    IF NOT "FRK_PersistImages".D003.Rows[8].Used OR "FRK_PersistImages".D003.Rows[8].SchemaVersion <> 4 OR "FRK_PersistImages".D003.Rows[8].ModelCode <> 'MODEL_B' OR "FRK_PersistImages".D003.Rows[8].Record.Scope <> 'StationA.Cell.Gate' OR "FRK_PersistImages".D003.Rows[8].Record.WriteKey <> 'preset' OR "FRK_PersistImages".D003.Rows[8].Record.Revision <> 2 OR "FRK_PersistImages".D003.Rows[8].Record.Kind <> 0 OR "FRK_PersistImages".D003.Rows[8].Record.ValueType <> 0 THEN RETURN; END_IF;
    #Ok := "FRK_ConfigDecode"(Text := STRING_TO_WSTRING("FRK_PersistImages".D003.Rows[8].Record.ValueText), Storage := 3, Minimum := 0.0, Maximum := 1000.0, MaxLength := 0, Value := "FRK_ConfigScratch".Value);
    IF NOT #Ok THEN RETURN; END_IF;
    IF NOT "FRK_PersistImages".D003.Rows[9].Used OR "FRK_PersistImages".D003.Rows[9].SchemaVersion <> 4 OR "FRK_PersistImages".D003.Rows[9].ModelCode <> 'MODEL_B' OR "FRK_PersistImages".D003.Rows[9].Record.Scope <> 'StationA.Satellite' OR "FRK_PersistImages".D003.Rows[9].Record.WriteKey <> 'timeout' OR "FRK_PersistImages".D003.Rows[9].Record.Revision <> 1 OR "FRK_PersistImages".D003.Rows[9].Record.Kind <> 0 OR "FRK_PersistImages".D003.Rows[9].Record.ValueType <> 3 THEN RETURN; END_IF;
    #Ok := "FRK_ConfigDecode"(Text := STRING_TO_WSTRING("FRK_PersistImages".D003.Rows[9].Record.ValueText), Storage := 7, Minimum := 1.0, Maximum := 60000.0, MaxLength := 0, Value := "FRK_ConfigScratch".Value);
    IF NOT #Ok THEN RETURN; END_IF;
    IF NOT "FRK_PersistImages".D003.Rows[10].Used OR "FRK_PersistImages".D003.Rows[10].SchemaVersion <> 4 OR "FRK_PersistImages".D003.Rows[10].ModelCode <> 'MODEL_B' OR "FRK_PersistImages".D003.Rows[10].Record.Scope <> 'StationA.Satellite' OR "FRK_PersistImages".D003.Rows[10].Record.WriteKey <> 'preset' OR "FRK_PersistImages".D003.Rows[10].Record.Revision <> 2 OR "FRK_PersistImages".D003.Rows[10].Record.Kind <> 0 OR "FRK_PersistImages".D003.Rows[10].Record.ValueType <> 0 THEN RETURN; END_IF;
    #Ok := "FRK_ConfigDecode"(Text := STRING_TO_WSTRING("FRK_PersistImages".D003.Rows[10].Record.ValueText), Storage := 3, Minimum := 0.0, Maximum := 1000.0, MaxLength := 0, Value := "FRK_ConfigScratch".Value);
    IF NOT #Ok THEN RETURN; END_IF;
    IF NOT "FRK_PersistImages".D003.Rows[11].Used OR "FRK_PersistImages".D003.Rows[11].SchemaVersion <> 4 OR "FRK_PersistImages".D003.Rows[11].ModelCode <> 'MODEL_B' OR "FRK_PersistImages".D003.Rows[11].Record.Scope <> 'StationA.Satellite.Cell' OR "FRK_PersistImages".D003.Rows[11].Record.WriteKey <> 'timeout' OR "FRK_PersistImages".D003.Rows[11].Record.Revision <> 1 OR "FRK_PersistImages".D003.Rows[11].Record.Kind <> 0 OR "FRK_PersistImages".D003.Rows[11].Record.ValueType <> 3 THEN RETURN; END_IF;
    #Ok := "FRK_ConfigDecode"(Text := STRING_TO_WSTRING("FRK_PersistImages".D003.Rows[11].Record.ValueText), Storage := 7, Minimum := 1.0, Maximum := 60000.0, MaxLength := 0, Value := "FRK_ConfigScratch".Value);
    IF NOT #Ok THEN RETURN; END_IF;
    IF NOT "FRK_PersistImages".D003.Rows[12].Used OR "FRK_PersistImages".D003.Rows[12].SchemaVersion <> 4 OR "FRK_PersistImages".D003.Rows[12].ModelCode <> 'MODEL_B' OR "FRK_PersistImages".D003.Rows[12].Record.Scope <> 'StationA.Satellite.Cell' OR "FRK_PersistImages".D003.Rows[12].Record.WriteKey <> 'preset' OR "FRK_PersistImages".D003.Rows[12].Record.Revision <> 2 OR "FRK_PersistImages".D003.Rows[12].Record.Kind <> 0 OR "FRK_PersistImages".D003.Rows[12].Record.ValueType <> 0 THEN RETURN; END_IF;
    #Ok := "FRK_ConfigDecode"(Text := STRING_TO_WSTRING("FRK_PersistImages".D003.Rows[12].Record.ValueText), Storage := 3, Minimum := 0.0, Maximum := 1000.0, MaxLength := 0, Value := "FRK_ConfigScratch".Value);
    IF NOT #Ok THEN RETURN; END_IF;
    IF NOT "FRK_PersistImages".D003.Rows[13].Used OR "FRK_PersistImages".D003.Rows[13].SchemaVersion <> 4 OR "FRK_PersistImages".D003.Rows[13].ModelCode <> 'MODEL_B' OR "FRK_PersistImages".D003.Rows[13].Record.Scope <> 'StationA.Satellite.Cell.Clamp' OR "FRK_PersistImages".D003.Rows[13].Record.WriteKey <> 'timeout' OR "FRK_PersistImages".D003.Rows[13].Record.Revision <> 1 OR "FRK_PersistImages".D003.Rows[13].Record.Kind <> 0 OR "FRK_PersistImages".D003.Rows[13].Record.ValueType <> 3 THEN RETURN; END_IF;
    #Ok := "FRK_ConfigDecode"(Text := STRING_TO_WSTRING("FRK_PersistImages".D003.Rows[13].Record.ValueText), Storage := 7, Minimum := 1.0, Maximum := 60000.0, MaxLength := 0, Value := "FRK_ConfigScratch".Value);
    IF NOT #Ok THEN RETURN; END_IF;
    IF NOT "FRK_PersistImages".D003.Rows[14].Used OR "FRK_PersistImages".D003.Rows[14].SchemaVersion <> 4 OR "FRK_PersistImages".D003.Rows[14].ModelCode <> 'MODEL_B' OR "FRK_PersistImages".D003.Rows[14].Record.Scope <> 'StationA.Satellite.Cell.Clamp' OR "FRK_PersistImages".D003.Rows[14].Record.WriteKey <> 'preset' OR "FRK_PersistImages".D003.Rows[14].Record.Revision <> 2 OR "FRK_PersistImages".D003.Rows[14].Record.Kind <> 0 OR "FRK_PersistImages".D003.Rows[14].Record.ValueType <> 0 THEN RETURN; END_IF;
    #Ok := "FRK_ConfigDecode"(Text := STRING_TO_WSTRING("FRK_PersistImages".D003.Rows[14].Record.ValueText), Storage := 3, Minimum := 0.0, Maximum := 1000.0, MaxLength := 0, Value := "FRK_ConfigScratch".Value);
    IF NOT #Ok THEN RETURN; END_IF;
    IF NOT "FRK_PersistImages".D003.Rows[15].Used OR "FRK_PersistImages".D003.Rows[15].SchemaVersion <> 4 OR "FRK_PersistImages".D003.Rows[15].ModelCode <> 'MODEL_B' OR "FRK_PersistImages".D003.Rows[15].Record.Scope <> 'StationA.Satellite.Cell.Gate' OR "FRK_PersistImages".D003.Rows[15].Record.WriteKey <> 'timeout' OR "FRK_PersistImages".D003.Rows[15].Record.Revision <> 1 OR "FRK_PersistImages".D003.Rows[15].Record.Kind <> 0 OR "FRK_PersistImages".D003.Rows[15].Record.ValueType <> 3 THEN RETURN; END_IF;
    #Ok := "FRK_ConfigDecode"(Text := STRING_TO_WSTRING("FRK_PersistImages".D003.Rows[15].Record.ValueText), Storage := 7, Minimum := 1.0, Maximum := 60000.0, MaxLength := 0, Value := "FRK_ConfigScratch".Value);
    IF NOT #Ok THEN RETURN; END_IF;
    IF NOT "FRK_PersistImages".D003.Rows[16].Used OR "FRK_PersistImages".D003.Rows[16].SchemaVersion <> 4 OR "FRK_PersistImages".D003.Rows[16].ModelCode <> 'MODEL_B' OR "FRK_PersistImages".D003.Rows[16].Record.Scope <> 'StationA.Satellite.Cell.Gate' OR "FRK_PersistImages".D003.Rows[16].Record.WriteKey <> 'preset' OR "FRK_PersistImages".D003.Rows[16].Record.Revision <> 2 OR "FRK_PersistImages".D003.Rows[16].Record.Kind <> 0 OR "FRK_PersistImages".D003.Rows[16].Record.ValueType <> 0 THEN RETURN; END_IF;
    #Ok := "FRK_ConfigDecode"(Text := STRING_TO_WSTRING("FRK_PersistImages".D003.Rows[16].Record.ValueText), Storage := 3, Minimum := 0.0, Maximum := 1000.0, MaxLength := 0, Value := "FRK_ConfigScratch".Value);
    IF NOT #Ok THEN RETURN; END_IF;
    IF NOT "FRK_PersistImages".D003.Rows[17].Used OR "FRK_PersistImages".D003.Rows[17].SchemaVersion <> 4 OR "FRK_PersistImages".D003.Rows[17].ModelCode <> 'MODEL_B' OR "FRK_PersistImages".D003.Rows[17].Record.Scope <> 'StationA.Satellite.Inner' OR "FRK_PersistImages".D003.Rows[17].Record.WriteKey <> 'timeout' OR "FRK_PersistImages".D003.Rows[17].Record.Revision <> 1 OR "FRK_PersistImages".D003.Rows[17].Record.Kind <> 0 OR "FRK_PersistImages".D003.Rows[17].Record.ValueType <> 3 THEN RETURN; END_IF;
    #Ok := "FRK_ConfigDecode"(Text := STRING_TO_WSTRING("FRK_PersistImages".D003.Rows[17].Record.ValueText), Storage := 7, Minimum := 1.0, Maximum := 60000.0, MaxLength := 0, Value := "FRK_ConfigScratch".Value);
    IF NOT #Ok THEN RETURN; END_IF;
    IF NOT "FRK_PersistImages".D003.Rows[18].Used OR "FRK_PersistImages".D003.Rows[18].SchemaVersion <> 4 OR "FRK_PersistImages".D003.Rows[18].ModelCode <> 'MODEL_B' OR "FRK_PersistImages".D003.Rows[18].Record.Scope <> 'StationA.Satellite.Inner' OR "FRK_PersistImages".D003.Rows[18].Record.WriteKey <> 'preset' OR "FRK_PersistImages".D003.Rows[18].Record.Revision <> 2 OR "FRK_PersistImages".D003.Rows[18].Record.Kind <> 0 OR "FRK_PersistImages".D003.Rows[18].Record.ValueType <> 0 THEN RETURN; END_IF;
    #Ok := "FRK_ConfigDecode"(Text := STRING_TO_WSTRING("FRK_PersistImages".D003.Rows[18].Record.ValueText), Storage := 3, Minimum := 0.0, Maximum := 1000.0, MaxLength := 0, Value := "FRK_ConfigScratch".Value);
    IF NOT #Ok THEN RETURN; END_IF;
    IF NOT "FRK_PersistImages".D003.Rows[19].Used OR "FRK_PersistImages".D003.Rows[19].SchemaVersion <> 4 OR "FRK_PersistImages".D003.Rows[19].ModelCode <> 'MODEL_B' OR "FRK_PersistImages".D003.Rows[19].Record.Scope <> 'StationA.Satellite.Inner.Cell' OR "FRK_PersistImages".D003.Rows[19].Record.WriteKey <> 'timeout' OR "FRK_PersistImages".D003.Rows[19].Record.Revision <> 1 OR "FRK_PersistImages".D003.Rows[19].Record.Kind <> 0 OR "FRK_PersistImages".D003.Rows[19].Record.ValueType <> 3 THEN RETURN; END_IF;
    #Ok := "FRK_ConfigDecode"(Text := STRING_TO_WSTRING("FRK_PersistImages".D003.Rows[19].Record.ValueText), Storage := 7, Minimum := 1.0, Maximum := 60000.0, MaxLength := 0, Value := "FRK_ConfigScratch".Value);
    IF NOT #Ok THEN RETURN; END_IF;
    IF NOT "FRK_PersistImages".D003.Rows[20].Used OR "FRK_PersistImages".D003.Rows[20].SchemaVersion <> 4 OR "FRK_PersistImages".D003.Rows[20].ModelCode <> 'MODEL_B' OR "FRK_PersistImages".D003.Rows[20].Record.Scope <> 'StationA.Satellite.Inner.Cell' OR "FRK_PersistImages".D003.Rows[20].Record.WriteKey <> 'preset' OR "FRK_PersistImages".D003.Rows[20].Record.Revision <> 2 OR "FRK_PersistImages".D003.Rows[20].Record.Kind <> 0 OR "FRK_PersistImages".D003.Rows[20].Record.ValueType <> 0 THEN RETURN; END_IF;
    #Ok := "FRK_ConfigDecode"(Text := STRING_TO_WSTRING("FRK_PersistImages".D003.Rows[20].Record.ValueText), Storage := 3, Minimum := 0.0, Maximum := 1000.0, MaxLength := 0, Value := "FRK_ConfigScratch".Value);
    IF NOT #Ok THEN RETURN; END_IF;
    IF NOT "FRK_PersistImages".D003.Rows[21].Used OR "FRK_PersistImages".D003.Rows[21].SchemaVersion <> 4 OR "FRK_PersistImages".D003.Rows[21].ModelCode <> 'MODEL_B' OR "FRK_PersistImages".D003.Rows[21].Record.Scope <> 'StationA.Satellite.Inner.Cell.Clamp' OR "FRK_PersistImages".D003.Rows[21].Record.WriteKey <> 'timeout' OR "FRK_PersistImages".D003.Rows[21].Record.Revision <> 1 OR "FRK_PersistImages".D003.Rows[21].Record.Kind <> 0 OR "FRK_PersistImages".D003.Rows[21].Record.ValueType <> 3 THEN RETURN; END_IF;
    #Ok := "FRK_ConfigDecode"(Text := STRING_TO_WSTRING("FRK_PersistImages".D003.Rows[21].Record.ValueText), Storage := 7, Minimum := 1.0, Maximum := 60000.0, MaxLength := 0, Value := "FRK_ConfigScratch".Value);
    IF NOT #Ok THEN RETURN; END_IF;
    IF NOT "FRK_PersistImages".D003.Rows[22].Used OR "FRK_PersistImages".D003.Rows[22].SchemaVersion <> 4 OR "FRK_PersistImages".D003.Rows[22].ModelCode <> 'MODEL_B' OR "FRK_PersistImages".D003.Rows[22].Record.Scope <> 'StationA.Satellite.Inner.Cell.Clamp' OR "FRK_PersistImages".D003.Rows[22].Record.WriteKey <> 'preset' OR "FRK_PersistImages".D003.Rows[22].Record.Revision <> 2 OR "FRK_PersistImages".D003.Rows[22].Record.Kind <> 0 OR "FRK_PersistImages".D003.Rows[22].Record.ValueType <> 0 THEN RETURN; END_IF;
    #Ok := "FRK_ConfigDecode"(Text := STRING_TO_WSTRING("FRK_PersistImages".D003.Rows[22].Record.ValueText), Storage := 3, Minimum := 0.0, Maximum := 1000.0, MaxLength := 0, Value := "FRK_ConfigScratch".Value);
    IF NOT #Ok THEN RETURN; END_IF;
    IF NOT "FRK_PersistImages".D003.Rows[23].Used OR "FRK_PersistImages".D003.Rows[23].SchemaVersion <> 4 OR "FRK_PersistImages".D003.Rows[23].ModelCode <> 'MODEL_B' OR "FRK_PersistImages".D003.Rows[23].Record.Scope <> 'StationA.Satellite.Inner.Cell.Gate' OR "FRK_PersistImages".D003.Rows[23].Record.WriteKey <> 'timeout' OR "FRK_PersistImages".D003.Rows[23].Record.Revision <> 1 OR "FRK_PersistImages".D003.Rows[23].Record.Kind <> 0 OR "FRK_PersistImages".D003.Rows[23].Record.ValueType <> 3 THEN RETURN; END_IF;
    #Ok := "FRK_ConfigDecode"(Text := STRING_TO_WSTRING("FRK_PersistImages".D003.Rows[23].Record.ValueText), Storage := 7, Minimum := 1.0, Maximum := 60000.0, MaxLength := 0, Value := "FRK_ConfigScratch".Value);
    IF NOT #Ok THEN RETURN; END_IF;
    IF NOT "FRK_PersistImages".D003.Rows[24].Used OR "FRK_PersistImages".D003.Rows[24].SchemaVersion <> 4 OR "FRK_PersistImages".D003.Rows[24].ModelCode <> 'MODEL_B' OR "FRK_PersistImages".D003.Rows[24].Record.Scope <> 'StationA.Satellite.Inner.Cell.Gate' OR "FRK_PersistImages".D003.Rows[24].Record.WriteKey <> 'preset' OR "FRK_PersistImages".D003.Rows[24].Record.Revision <> 2 OR "FRK_PersistImages".D003.Rows[24].Record.Kind <> 0 OR "FRK_PersistImages".D003.Rows[24].Record.ValueType <> 0 THEN RETURN; END_IF;
    #Ok := "FRK_ConfigDecode"(Text := STRING_TO_WSTRING("FRK_PersistImages".D003.Rows[24].Record.ValueText), Storage := 3, Minimum := 0.0, Maximum := 1000.0, MaxLength := 0, Value := "FRK_ConfigScratch".Value);
    IF NOT #Ok THEN RETURN; END_IF;
    #Stored := "FRK_ConfigFind"(Scope := 'StationA', Key := 'timeout', ModelCode := 'MODEL_B');
    IF #Stored = 0 THEN
        FOR #Stored := 1 TO 108 DO IF NOT "FRK_ConfigStore".Rows[#Stored].Used THEN EXIT; END_IF; END_FOR;
    END_IF;
    IF #Stored < 1 OR #Stored > 108 THEN RETURN; END_IF;
    "FRK_ConfigStore".Rows[#Stored] := "FRK_PersistImages".D003.Rows[1];
    #Stored := "FRK_ConfigFind"(Scope := 'StationA', Key := 'preset', ModelCode := 'MODEL_B');
    IF #Stored = 0 THEN
        FOR #Stored := 1 TO 108 DO IF NOT "FRK_ConfigStore".Rows[#Stored].Used THEN EXIT; END_IF; END_FOR;
    END_IF;
    IF #Stored < 1 OR #Stored > 108 THEN RETURN; END_IF;
    "FRK_ConfigStore".Rows[#Stored] := "FRK_PersistImages".D003.Rows[2];
    #Stored := "FRK_ConfigFind"(Scope := 'StationA.Cell', Key := 'timeout', ModelCode := 'MODEL_B');
    IF #Stored = 0 THEN
        FOR #Stored := 1 TO 108 DO IF NOT "FRK_ConfigStore".Rows[#Stored].Used THEN EXIT; END_IF; END_FOR;
    END_IF;
    IF #Stored < 1 OR #Stored > 108 THEN RETURN; END_IF;
    "FRK_ConfigStore".Rows[#Stored] := "FRK_PersistImages".D003.Rows[3];
    #Stored := "FRK_ConfigFind"(Scope := 'StationA.Cell', Key := 'preset', ModelCode := 'MODEL_B');
    IF #Stored = 0 THEN
        FOR #Stored := 1 TO 108 DO IF NOT "FRK_ConfigStore".Rows[#Stored].Used THEN EXIT; END_IF; END_FOR;
    END_IF;
    IF #Stored < 1 OR #Stored > 108 THEN RETURN; END_IF;
    "FRK_ConfigStore".Rows[#Stored] := "FRK_PersistImages".D003.Rows[4];
    #Stored := "FRK_ConfigFind"(Scope := 'StationA.Cell.Clamp', Key := 'timeout', ModelCode := 'MODEL_B');
    IF #Stored = 0 THEN
        FOR #Stored := 1 TO 108 DO IF NOT "FRK_ConfigStore".Rows[#Stored].Used THEN EXIT; END_IF; END_FOR;
    END_IF;
    IF #Stored < 1 OR #Stored > 108 THEN RETURN; END_IF;
    "FRK_ConfigStore".Rows[#Stored] := "FRK_PersistImages".D003.Rows[5];
    #Stored := "FRK_ConfigFind"(Scope := 'StationA.Cell.Clamp', Key := 'preset', ModelCode := 'MODEL_B');
    IF #Stored = 0 THEN
        FOR #Stored := 1 TO 108 DO IF NOT "FRK_ConfigStore".Rows[#Stored].Used THEN EXIT; END_IF; END_FOR;
    END_IF;
    IF #Stored < 1 OR #Stored > 108 THEN RETURN; END_IF;
    "FRK_ConfigStore".Rows[#Stored] := "FRK_PersistImages".D003.Rows[6];
    #Stored := "FRK_ConfigFind"(Scope := 'StationA.Cell.Gate', Key := 'timeout', ModelCode := 'MODEL_B');
    IF #Stored = 0 THEN
        FOR #Stored := 1 TO 108 DO IF NOT "FRK_ConfigStore".Rows[#Stored].Used THEN EXIT; END_IF; END_FOR;
    END_IF;
    IF #Stored < 1 OR #Stored > 108 THEN RETURN; END_IF;
    "FRK_ConfigStore".Rows[#Stored] := "FRK_PersistImages".D003.Rows[7];
    #Stored := "FRK_ConfigFind"(Scope := 'StationA.Cell.Gate', Key := 'preset', ModelCode := 'MODEL_B');
    IF #Stored = 0 THEN
        FOR #Stored := 1 TO 108 DO IF NOT "FRK_ConfigStore".Rows[#Stored].Used THEN EXIT; END_IF; END_FOR;
    END_IF;
    IF #Stored < 1 OR #Stored > 108 THEN RETURN; END_IF;
    "FRK_ConfigStore".Rows[#Stored] := "FRK_PersistImages".D003.Rows[8];
    #Stored := "FRK_ConfigFind"(Scope := 'StationA.Satellite', Key := 'timeout', ModelCode := 'MODEL_B');
    IF #Stored = 0 THEN
        FOR #Stored := 1 TO 108 DO IF NOT "FRK_ConfigStore".Rows[#Stored].Used THEN EXIT; END_IF; END_FOR;
    END_IF;
    IF #Stored < 1 OR #Stored > 108 THEN RETURN; END_IF;
    "FRK_ConfigStore".Rows[#Stored] := "FRK_PersistImages".D003.Rows[9];
    #Stored := "FRK_ConfigFind"(Scope := 'StationA.Satellite', Key := 'preset', ModelCode := 'MODEL_B');
    IF #Stored = 0 THEN
        FOR #Stored := 1 TO 108 DO IF NOT "FRK_ConfigStore".Rows[#Stored].Used THEN EXIT; END_IF; END_FOR;
    END_IF;
    IF #Stored < 1 OR #Stored > 108 THEN RETURN; END_IF;
    "FRK_ConfigStore".Rows[#Stored] := "FRK_PersistImages".D003.Rows[10];
    #Stored := "FRK_ConfigFind"(Scope := 'StationA.Satellite.Cell', Key := 'timeout', ModelCode := 'MODEL_B');
    IF #Stored = 0 THEN
        FOR #Stored := 1 TO 108 DO IF NOT "FRK_ConfigStore".Rows[#Stored].Used THEN EXIT; END_IF; END_FOR;
    END_IF;
    IF #Stored < 1 OR #Stored > 108 THEN RETURN; END_IF;
    "FRK_ConfigStore".Rows[#Stored] := "FRK_PersistImages".D003.Rows[11];
    #Stored := "FRK_ConfigFind"(Scope := 'StationA.Satellite.Cell', Key := 'preset', ModelCode := 'MODEL_B');
    IF #Stored = 0 THEN
        FOR #Stored := 1 TO 108 DO IF NOT "FRK_ConfigStore".Rows[#Stored].Used THEN EXIT; END_IF; END_FOR;
    END_IF;
    IF #Stored < 1 OR #Stored > 108 THEN RETURN; END_IF;
    "FRK_ConfigStore".Rows[#Stored] := "FRK_PersistImages".D003.Rows[12];
    #Stored := "FRK_ConfigFind"(Scope := 'StationA.Satellite.Cell.Clamp', Key := 'timeout', ModelCode := 'MODEL_B');
    IF #Stored = 0 THEN
        FOR #Stored := 1 TO 108 DO IF NOT "FRK_ConfigStore".Rows[#Stored].Used THEN EXIT; END_IF; END_FOR;
    END_IF;
    IF #Stored < 1 OR #Stored > 108 THEN RETURN; END_IF;
    "FRK_ConfigStore".Rows[#Stored] := "FRK_PersistImages".D003.Rows[13];
    #Stored := "FRK_ConfigFind"(Scope := 'StationA.Satellite.Cell.Clamp', Key := 'preset', ModelCode := 'MODEL_B');
    IF #Stored = 0 THEN
        FOR #Stored := 1 TO 108 DO IF NOT "FRK_ConfigStore".Rows[#Stored].Used THEN EXIT; END_IF; END_FOR;
    END_IF;
    IF #Stored < 1 OR #Stored > 108 THEN RETURN; END_IF;
    "FRK_ConfigStore".Rows[#Stored] := "FRK_PersistImages".D003.Rows[14];
    #Stored := "FRK_ConfigFind"(Scope := 'StationA.Satellite.Cell.Gate', Key := 'timeout', ModelCode := 'MODEL_B');
    IF #Stored = 0 THEN
        FOR #Stored := 1 TO 108 DO IF NOT "FRK_ConfigStore".Rows[#Stored].Used THEN EXIT; END_IF; END_FOR;
    END_IF;
    IF #Stored < 1 OR #Stored > 108 THEN RETURN; END_IF;
    "FRK_ConfigStore".Rows[#Stored] := "FRK_PersistImages".D003.Rows[15];
    #Stored := "FRK_ConfigFind"(Scope := 'StationA.Satellite.Cell.Gate', Key := 'preset', ModelCode := 'MODEL_B');
    IF #Stored = 0 THEN
        FOR #Stored := 1 TO 108 DO IF NOT "FRK_ConfigStore".Rows[#Stored].Used THEN EXIT; END_IF; END_FOR;
    END_IF;
    IF #Stored < 1 OR #Stored > 108 THEN RETURN; END_IF;
    "FRK_ConfigStore".Rows[#Stored] := "FRK_PersistImages".D003.Rows[16];
    #Stored := "FRK_ConfigFind"(Scope := 'StationA.Satellite.Inner', Key := 'timeout', ModelCode := 'MODEL_B');
    IF #Stored = 0 THEN
        FOR #Stored := 1 TO 108 DO IF NOT "FRK_ConfigStore".Rows[#Stored].Used THEN EXIT; END_IF; END_FOR;
    END_IF;
    IF #Stored < 1 OR #Stored > 108 THEN RETURN; END_IF;
    "FRK_ConfigStore".Rows[#Stored] := "FRK_PersistImages".D003.Rows[17];
    #Stored := "FRK_ConfigFind"(Scope := 'StationA.Satellite.Inner', Key := 'preset', ModelCode := 'MODEL_B');
    IF #Stored = 0 THEN
        FOR #Stored := 1 TO 108 DO IF NOT "FRK_ConfigStore".Rows[#Stored].Used THEN EXIT; END_IF; END_FOR;
    END_IF;
    IF #Stored < 1 OR #Stored > 108 THEN RETURN; END_IF;
    "FRK_ConfigStore".Rows[#Stored] := "FRK_PersistImages".D003.Rows[18];
    #Stored := "FRK_ConfigFind"(Scope := 'StationA.Satellite.Inner.Cell', Key := 'timeout', ModelCode := 'MODEL_B');
    IF #Stored = 0 THEN
        FOR #Stored := 1 TO 108 DO IF NOT "FRK_ConfigStore".Rows[#Stored].Used THEN EXIT; END_IF; END_FOR;
    END_IF;
    IF #Stored < 1 OR #Stored > 108 THEN RETURN; END_IF;
    "FRK_ConfigStore".Rows[#Stored] := "FRK_PersistImages".D003.Rows[19];
    #Stored := "FRK_ConfigFind"(Scope := 'StationA.Satellite.Inner.Cell', Key := 'preset', ModelCode := 'MODEL_B');
    IF #Stored = 0 THEN
        FOR #Stored := 1 TO 108 DO IF NOT "FRK_ConfigStore".Rows[#Stored].Used THEN EXIT; END_IF; END_FOR;
    END_IF;
    IF #Stored < 1 OR #Stored > 108 THEN RETURN; END_IF;
    "FRK_ConfigStore".Rows[#Stored] := "FRK_PersistImages".D003.Rows[20];
    #Stored := "FRK_ConfigFind"(Scope := 'StationA.Satellite.Inner.Cell.Clamp', Key := 'timeout', ModelCode := 'MODEL_B');
    IF #Stored = 0 THEN
        FOR #Stored := 1 TO 108 DO IF NOT "FRK_ConfigStore".Rows[#Stored].Used THEN EXIT; END_IF; END_FOR;
    END_IF;
    IF #Stored < 1 OR #Stored > 108 THEN RETURN; END_IF;
    "FRK_ConfigStore".Rows[#Stored] := "FRK_PersistImages".D003.Rows[21];
    #Stored := "FRK_ConfigFind"(Scope := 'StationA.Satellite.Inner.Cell.Clamp', Key := 'preset', ModelCode := 'MODEL_B');
    IF #Stored = 0 THEN
        FOR #Stored := 1 TO 108 DO IF NOT "FRK_ConfigStore".Rows[#Stored].Used THEN EXIT; END_IF; END_FOR;
    END_IF;
    IF #Stored < 1 OR #Stored > 108 THEN RETURN; END_IF;
    "FRK_ConfigStore".Rows[#Stored] := "FRK_PersistImages".D003.Rows[22];
    #Stored := "FRK_ConfigFind"(Scope := 'StationA.Satellite.Inner.Cell.Gate', Key := 'timeout', ModelCode := 'MODEL_B');
    IF #Stored = 0 THEN
        FOR #Stored := 1 TO 108 DO IF NOT "FRK_ConfigStore".Rows[#Stored].Used THEN EXIT; END_IF; END_FOR;
    END_IF;
    IF #Stored < 1 OR #Stored > 108 THEN RETURN; END_IF;
    "FRK_ConfigStore".Rows[#Stored] := "FRK_PersistImages".D003.Rows[23];
    #Stored := "FRK_ConfigFind"(Scope := 'StationA.Satellite.Inner.Cell.Gate', Key := 'preset', ModelCode := 'MODEL_B');
    IF #Stored = 0 THEN
        FOR #Stored := 1 TO 108 DO IF NOT "FRK_ConfigStore".Rows[#Stored].Used THEN EXIT; END_IF; END_FOR;
    END_IF;
    IF #Stored < 1 OR #Stored > 108 THEN RETURN; END_IF;
    "FRK_ConfigStore".Rows[#Stored] := "FRK_PersistImages".D003.Rows[24];
    "FRK_ConfigStore".SchemaVersion := 1;
    #FRK_DocApply_D003 := TRUE;
END_FUNCTION
FUNCTION "FRK_DocCapture_D004" : Bool
{ S7_Optimized_Access := 'TRUE' }
VERSION : 0.1
VAR_IN_OUT
    Length : DInt;
END_VAR
VAR_TEMP
    Index : Int;
    Stored : Int;
    Position : DInt;
    NativeResult : Int;
    Ok : Bool;
END_VAR
BEGIN
    #FRK_DocCapture_D004 := FALSE;
    "FRK_PersistImages".D004.SchemaVersion := 1; "FRK_PersistImages".D004.Scope := 'StationA';
    #Stored := 0;
    FOR #Index := 1 TO 2 DO
        IF "FRK_AccessPolicies".Rows[#Index].Scope = 'StationA' THEN #Stored := #Index; END_IF;
    END_FOR;
    IF #Stored = 0 THEN RETURN; END_IF;
    "FRK_PersistImages".D004.Image := "FRK_AccessPolicies".Rows[#Stored];
    IF NOT "FRK_AccessPolicyValid"(Image := "FRK_PersistImages".D004.Image) THEN RETURN; END_IF;
    FOR #Index := 0 TO 413 DO "FRK_PersistBuffers".D004Data[#Index] := BYTE#0; END_FOR;
    #Position := 24;
    #NativeResult := Serialize(SRC_VARIABLE := "FRK_PersistImages".D004, DEST_ARRAY => "FRK_PersistBuffers".D004Data, POS := #Position);
    IF #NativeResult <> 0 OR #Position < 24 OR #Position > 414 THEN RETURN; END_IF;
    #Length := #Position - 24;
    #FRK_DocCapture_D004 := TRUE;
END_FUNCTION
FUNCTION "FRK_DocApply_D004" : Bool
{ S7_Optimized_Access := 'TRUE' }
VERSION : 0.1
VAR_TEMP
    Index : Int;
    Stored : Int;
    Position : DInt;
    NativeResult : Int;
    Ok : Bool;
END_VAR
BEGIN
    #FRK_DocApply_D004 := FALSE;
    #Position := 24;
    #NativeResult := Deserialize(SRC_ARRAY := "FRK_PersistBuffers".D004Data, DEST_VARIABLE => "FRK_PersistImages".D004, POS := #Position);
    IF #NativeResult <> 0 OR #Position <> 24 + UDINT_TO_DINT("FRK_PersistConsumers".Rows[4].Result.Length) THEN RETURN; END_IF;
    IF "FRK_PersistImages".D004.SchemaVersion <> 1 OR "FRK_PersistImages".D004.Scope <> 'StationA' THEN RETURN; END_IF;
    IF "FRK_PersistImages".D004.Image.Scope <> 'StationA' OR NOT "FRK_AccessPolicyValid"(Image := "FRK_PersistImages".D004.Image) THEN RETURN; END_IF;
    "FRK_AccessPolicies".Rows[1] := "FRK_PersistImages".D004.Image;
    #FRK_DocApply_D004 := TRUE;
END_FUNCTION
FUNCTION "FRK_DocCapture_D005" : Bool
{ S7_Optimized_Access := 'TRUE' }
VERSION : 0.1
VAR_IN_OUT
    Length : DInt;
END_VAR
VAR_TEMP
    Index : Int;
    Stored : Int;
    Position : DInt;
    NativeResult : Int;
    Ok : Bool;
END_VAR
BEGIN
    #FRK_DocCapture_D005 := FALSE;
    "FRK_PersistImages".D005.SchemaVersion := 1; "FRK_PersistImages".D005.Scope := 'StationB';
    "FRK_PersistImages".D005.Kind := 1;
    "FRK_PersistImages".D005.ModelCode := '';
    "FRK_PersistImages".D005.ActiveModel := "FRK_ConfigStore".ActiveModels[2];
    "FRK_PersistImages".D005.Count := 6;
    #Stored := "FRK_ConfigFind"(Scope := 'StationB', Key := 'siteLabel', ModelCode := '');
    IF #Stored = 0 THEN RETURN; END_IF;
    "FRK_PersistImages".D005.Rows[1] := "FRK_ConfigStore".Rows[#Stored];
    #Stored := "FRK_ConfigFind"(Scope := 'StationB', Key := 'enabled', ModelCode := '');
    IF #Stored = 0 THEN RETURN; END_IF;
    "FRK_PersistImages".D005.Rows[2] := "FRK_ConfigStore".Rows[#Stored];
    #Stored := "FRK_ConfigFind"(Scope := 'StationB.Satellite', Key := 'siteLabel', ModelCode := '');
    IF #Stored = 0 THEN RETURN; END_IF;
    "FRK_PersistImages".D005.Rows[3] := "FRK_ConfigStore".Rows[#Stored];
    #Stored := "FRK_ConfigFind"(Scope := 'StationB.Satellite', Key := 'enabled', ModelCode := '');
    IF #Stored = 0 THEN RETURN; END_IF;
    "FRK_PersistImages".D005.Rows[4] := "FRK_ConfigStore".Rows[#Stored];
    #Stored := "FRK_ConfigFind"(Scope := 'StationB.Satellite.Inner', Key := 'siteLabel', ModelCode := '');
    IF #Stored = 0 THEN RETURN; END_IF;
    "FRK_PersistImages".D005.Rows[5] := "FRK_ConfigStore".Rows[#Stored];
    #Stored := "FRK_ConfigFind"(Scope := 'StationB.Satellite.Inner', Key := 'enabled', ModelCode := '');
    IF #Stored = 0 THEN RETURN; END_IF;
    "FRK_PersistImages".D005.Rows[6] := "FRK_ConfigStore".Rows[#Stored];
    FOR #Index := 0 TO 3085 DO "FRK_PersistBuffers".D005Data[#Index] := BYTE#0; END_FOR;
    #Position := 24;
    #NativeResult := Serialize(SRC_VARIABLE := "FRK_PersistImages".D005, DEST_ARRAY => "FRK_PersistBuffers".D005Data, POS := #Position);
    IF #NativeResult <> 0 OR #Position < 24 OR #Position > 3086 THEN RETURN; END_IF;
    #Length := #Position - 24;
    #FRK_DocCapture_D005 := TRUE;
END_FUNCTION
FUNCTION "FRK_DocApply_D005" : Bool
{ S7_Optimized_Access := 'TRUE' }
VERSION : 0.1
VAR_TEMP
    Index : Int;
    Stored : Int;
    Position : DInt;
    NativeResult : Int;
    Ok : Bool;
END_VAR
BEGIN
    #FRK_DocApply_D005 := FALSE;
    #Position := 24;
    #NativeResult := Deserialize(SRC_ARRAY := "FRK_PersistBuffers".D005Data, DEST_VARIABLE => "FRK_PersistImages".D005, POS := #Position);
    IF #NativeResult <> 0 OR #Position <> 24 + UDINT_TO_DINT("FRK_PersistConsumers".Rows[5].Result.Length) THEN RETURN; END_IF;
    IF "FRK_PersistImages".D005.SchemaVersion <> 1 OR "FRK_PersistImages".D005.Scope <> 'StationB' THEN RETURN; END_IF;
    IF "FRK_PersistImages".D005.Kind <> 1 OR "FRK_PersistImages".D005.ModelCode <> '' OR "FRK_PersistImages".D005.Count <> 6 THEN RETURN; END_IF;
    IF "FRK_PersistImages".D005.ActiveModel <> 'MODEL_A' AND "FRK_PersistImages".D005.ActiveModel <> 'MODEL_B' THEN RETURN; END_IF;
    IF NOT "FRK_PersistImages".D005.Rows[1].Used OR "FRK_PersistImages".D005.Rows[1].SchemaVersion <> 1 OR "FRK_PersistImages".D005.Rows[1].ModelCode <> '' OR "FRK_PersistImages".D005.Rows[1].Record.Scope <> 'StationB' OR "FRK_PersistImages".D005.Rows[1].Record.WriteKey <> 'siteLabel' OR "FRK_PersistImages".D005.Rows[1].Record.Revision <> 1 OR "FRK_PersistImages".D005.Rows[1].Record.Kind <> 1 OR "FRK_PersistImages".D005.Rows[1].Record.ValueType <> 1 THEN RETURN; END_IF;
    #Ok := "FRK_ConfigDecode"(Text := STRING_TO_WSTRING("FRK_PersistImages".D005.Rows[1].Record.ValueText), Storage := 8, Minimum := 0.0, Maximum := 1.0, MaxLength := 80, Value := "FRK_ConfigScratch".Value);
    IF NOT #Ok THEN RETURN; END_IF;
    IF NOT "FRK_PersistImages".D005.Rows[2].Used OR "FRK_PersistImages".D005.Rows[2].SchemaVersion <> 1 OR "FRK_PersistImages".D005.Rows[2].ModelCode <> '' OR "FRK_PersistImages".D005.Rows[2].Record.Scope <> 'StationB' OR "FRK_PersistImages".D005.Rows[2].Record.WriteKey <> 'enabled' OR "FRK_PersistImages".D005.Rows[2].Record.Revision <> 1 OR "FRK_PersistImages".D005.Rows[2].Record.Kind <> 1 OR "FRK_PersistImages".D005.Rows[2].Record.ValueType <> 2 THEN RETURN; END_IF;
    #Ok := "FRK_ConfigDecode"(Text := STRING_TO_WSTRING("FRK_PersistImages".D005.Rows[2].Record.ValueText), Storage := 1, Minimum := 0.0, Maximum := 1.0, MaxLength := 0, Value := "FRK_ConfigScratch".Value);
    IF NOT #Ok THEN RETURN; END_IF;
    IF NOT "FRK_PersistImages".D005.Rows[3].Used OR "FRK_PersistImages".D005.Rows[3].SchemaVersion <> 1 OR "FRK_PersistImages".D005.Rows[3].ModelCode <> '' OR "FRK_PersistImages".D005.Rows[3].Record.Scope <> 'StationB.Satellite' OR "FRK_PersistImages".D005.Rows[3].Record.WriteKey <> 'siteLabel' OR "FRK_PersistImages".D005.Rows[3].Record.Revision <> 1 OR "FRK_PersistImages".D005.Rows[3].Record.Kind <> 1 OR "FRK_PersistImages".D005.Rows[3].Record.ValueType <> 1 THEN RETURN; END_IF;
    #Ok := "FRK_ConfigDecode"(Text := STRING_TO_WSTRING("FRK_PersistImages".D005.Rows[3].Record.ValueText), Storage := 8, Minimum := 0.0, Maximum := 1.0, MaxLength := 80, Value := "FRK_ConfigScratch".Value);
    IF NOT #Ok THEN RETURN; END_IF;
    IF NOT "FRK_PersistImages".D005.Rows[4].Used OR "FRK_PersistImages".D005.Rows[4].SchemaVersion <> 1 OR "FRK_PersistImages".D005.Rows[4].ModelCode <> '' OR "FRK_PersistImages".D005.Rows[4].Record.Scope <> 'StationB.Satellite' OR "FRK_PersistImages".D005.Rows[4].Record.WriteKey <> 'enabled' OR "FRK_PersistImages".D005.Rows[4].Record.Revision <> 1 OR "FRK_PersistImages".D005.Rows[4].Record.Kind <> 1 OR "FRK_PersistImages".D005.Rows[4].Record.ValueType <> 2 THEN RETURN; END_IF;
    #Ok := "FRK_ConfigDecode"(Text := STRING_TO_WSTRING("FRK_PersistImages".D005.Rows[4].Record.ValueText), Storage := 1, Minimum := 0.0, Maximum := 1.0, MaxLength := 0, Value := "FRK_ConfigScratch".Value);
    IF NOT #Ok THEN RETURN; END_IF;
    IF NOT "FRK_PersistImages".D005.Rows[5].Used OR "FRK_PersistImages".D005.Rows[5].SchemaVersion <> 1 OR "FRK_PersistImages".D005.Rows[5].ModelCode <> '' OR "FRK_PersistImages".D005.Rows[5].Record.Scope <> 'StationB.Satellite.Inner' OR "FRK_PersistImages".D005.Rows[5].Record.WriteKey <> 'siteLabel' OR "FRK_PersistImages".D005.Rows[5].Record.Revision <> 1 OR "FRK_PersistImages".D005.Rows[5].Record.Kind <> 1 OR "FRK_PersistImages".D005.Rows[5].Record.ValueType <> 1 THEN RETURN; END_IF;
    #Ok := "FRK_ConfigDecode"(Text := STRING_TO_WSTRING("FRK_PersistImages".D005.Rows[5].Record.ValueText), Storage := 8, Minimum := 0.0, Maximum := 1.0, MaxLength := 80, Value := "FRK_ConfigScratch".Value);
    IF NOT #Ok THEN RETURN; END_IF;
    IF NOT "FRK_PersistImages".D005.Rows[6].Used OR "FRK_PersistImages".D005.Rows[6].SchemaVersion <> 1 OR "FRK_PersistImages".D005.Rows[6].ModelCode <> '' OR "FRK_PersistImages".D005.Rows[6].Record.Scope <> 'StationB.Satellite.Inner' OR "FRK_PersistImages".D005.Rows[6].Record.WriteKey <> 'enabled' OR "FRK_PersistImages".D005.Rows[6].Record.Revision <> 1 OR "FRK_PersistImages".D005.Rows[6].Record.Kind <> 1 OR "FRK_PersistImages".D005.Rows[6].Record.ValueType <> 2 THEN RETURN; END_IF;
    #Ok := "FRK_ConfigDecode"(Text := STRING_TO_WSTRING("FRK_PersistImages".D005.Rows[6].Record.ValueText), Storage := 1, Minimum := 0.0, Maximum := 1.0, MaxLength := 0, Value := "FRK_ConfigScratch".Value);
    IF NOT #Ok THEN RETURN; END_IF;
    #Stored := "FRK_ConfigFind"(Scope := 'StationB', Key := 'siteLabel', ModelCode := '');
    IF #Stored = 0 THEN
        FOR #Stored := 1 TO 108 DO IF NOT "FRK_ConfigStore".Rows[#Stored].Used THEN EXIT; END_IF; END_FOR;
    END_IF;
    IF #Stored < 1 OR #Stored > 108 THEN RETURN; END_IF;
    "FRK_ConfigStore".Rows[#Stored] := "FRK_PersistImages".D005.Rows[1];
    #Stored := "FRK_ConfigFind"(Scope := 'StationB', Key := 'enabled', ModelCode := '');
    IF #Stored = 0 THEN
        FOR #Stored := 1 TO 108 DO IF NOT "FRK_ConfigStore".Rows[#Stored].Used THEN EXIT; END_IF; END_FOR;
    END_IF;
    IF #Stored < 1 OR #Stored > 108 THEN RETURN; END_IF;
    "FRK_ConfigStore".Rows[#Stored] := "FRK_PersistImages".D005.Rows[2];
    #Stored := "FRK_ConfigFind"(Scope := 'StationB.Satellite', Key := 'siteLabel', ModelCode := '');
    IF #Stored = 0 THEN
        FOR #Stored := 1 TO 108 DO IF NOT "FRK_ConfigStore".Rows[#Stored].Used THEN EXIT; END_IF; END_FOR;
    END_IF;
    IF #Stored < 1 OR #Stored > 108 THEN RETURN; END_IF;
    "FRK_ConfigStore".Rows[#Stored] := "FRK_PersistImages".D005.Rows[3];
    #Stored := "FRK_ConfigFind"(Scope := 'StationB.Satellite', Key := 'enabled', ModelCode := '');
    IF #Stored = 0 THEN
        FOR #Stored := 1 TO 108 DO IF NOT "FRK_ConfigStore".Rows[#Stored].Used THEN EXIT; END_IF; END_FOR;
    END_IF;
    IF #Stored < 1 OR #Stored > 108 THEN RETURN; END_IF;
    "FRK_ConfigStore".Rows[#Stored] := "FRK_PersistImages".D005.Rows[4];
    #Stored := "FRK_ConfigFind"(Scope := 'StationB.Satellite.Inner', Key := 'siteLabel', ModelCode := '');
    IF #Stored = 0 THEN
        FOR #Stored := 1 TO 108 DO IF NOT "FRK_ConfigStore".Rows[#Stored].Used THEN EXIT; END_IF; END_FOR;
    END_IF;
    IF #Stored < 1 OR #Stored > 108 THEN RETURN; END_IF;
    "FRK_ConfigStore".Rows[#Stored] := "FRK_PersistImages".D005.Rows[5];
    #Stored := "FRK_ConfigFind"(Scope := 'StationB.Satellite.Inner', Key := 'enabled', ModelCode := '');
    IF #Stored = 0 THEN
        FOR #Stored := 1 TO 108 DO IF NOT "FRK_ConfigStore".Rows[#Stored].Used THEN EXIT; END_IF; END_FOR;
    END_IF;
    IF #Stored < 1 OR #Stored > 108 THEN RETURN; END_IF;
    "FRK_ConfigStore".Rows[#Stored] := "FRK_PersistImages".D005.Rows[6];
    "FRK_ConfigStore".ActiveModels[2] := "FRK_PersistImages".D005.ActiveModel;
    "FRK_ConfigStore".SchemaVersion := 1;
    #FRK_DocApply_D005 := TRUE;
END_FUNCTION
FUNCTION "FRK_DocCapture_D006" : Bool
{ S7_Optimized_Access := 'TRUE' }
VERSION : 0.1
VAR_IN_OUT
    Length : DInt;
END_VAR
VAR_TEMP
    Index : Int;
    Stored : Int;
    Position : DInt;
    NativeResult : Int;
    Ok : Bool;
END_VAR
BEGIN
    #FRK_DocCapture_D006 := FALSE;
    "FRK_PersistImages".D006.SchemaVersion := 1; "FRK_PersistImages".D006.Scope := 'StationB';
    "FRK_PersistImages".D006.Kind := 0;
    "FRK_PersistImages".D006.ModelCode := 'MODEL_A';
    "FRK_PersistImages".D006.ActiveModel := "FRK_ConfigStore".ActiveModels[2];
    "FRK_PersistImages".D006.Count := 24;
    #Stored := "FRK_ConfigFind"(Scope := 'StationB', Key := 'timeout', ModelCode := 'MODEL_A');
    IF #Stored = 0 THEN RETURN; END_IF;
    "FRK_PersistImages".D006.Rows[1] := "FRK_ConfigStore".Rows[#Stored];
    #Stored := "FRK_ConfigFind"(Scope := 'StationB', Key := 'preset', ModelCode := 'MODEL_A');
    IF #Stored = 0 THEN RETURN; END_IF;
    "FRK_PersistImages".D006.Rows[2] := "FRK_ConfigStore".Rows[#Stored];
    #Stored := "FRK_ConfigFind"(Scope := 'StationB.Cell', Key := 'timeout', ModelCode := 'MODEL_A');
    IF #Stored = 0 THEN RETURN; END_IF;
    "FRK_PersistImages".D006.Rows[3] := "FRK_ConfigStore".Rows[#Stored];
    #Stored := "FRK_ConfigFind"(Scope := 'StationB.Cell', Key := 'preset', ModelCode := 'MODEL_A');
    IF #Stored = 0 THEN RETURN; END_IF;
    "FRK_PersistImages".D006.Rows[4] := "FRK_ConfigStore".Rows[#Stored];
    #Stored := "FRK_ConfigFind"(Scope := 'StationB.Cell.Clamp', Key := 'timeout', ModelCode := 'MODEL_A');
    IF #Stored = 0 THEN RETURN; END_IF;
    "FRK_PersistImages".D006.Rows[5] := "FRK_ConfigStore".Rows[#Stored];
    #Stored := "FRK_ConfigFind"(Scope := 'StationB.Cell.Clamp', Key := 'preset', ModelCode := 'MODEL_A');
    IF #Stored = 0 THEN RETURN; END_IF;
    "FRK_PersistImages".D006.Rows[6] := "FRK_ConfigStore".Rows[#Stored];
    #Stored := "FRK_ConfigFind"(Scope := 'StationB.Cell.Gate', Key := 'timeout', ModelCode := 'MODEL_A');
    IF #Stored = 0 THEN RETURN; END_IF;
    "FRK_PersistImages".D006.Rows[7] := "FRK_ConfigStore".Rows[#Stored];
    #Stored := "FRK_ConfigFind"(Scope := 'StationB.Cell.Gate', Key := 'preset', ModelCode := 'MODEL_A');
    IF #Stored = 0 THEN RETURN; END_IF;
    "FRK_PersistImages".D006.Rows[8] := "FRK_ConfigStore".Rows[#Stored];
    #Stored := "FRK_ConfigFind"(Scope := 'StationB.Satellite', Key := 'timeout', ModelCode := 'MODEL_A');
    IF #Stored = 0 THEN RETURN; END_IF;
    "FRK_PersistImages".D006.Rows[9] := "FRK_ConfigStore".Rows[#Stored];
    #Stored := "FRK_ConfigFind"(Scope := 'StationB.Satellite', Key := 'preset', ModelCode := 'MODEL_A');
    IF #Stored = 0 THEN RETURN; END_IF;
    "FRK_PersistImages".D006.Rows[10] := "FRK_ConfigStore".Rows[#Stored];
    #Stored := "FRK_ConfigFind"(Scope := 'StationB.Satellite.Cell', Key := 'timeout', ModelCode := 'MODEL_A');
    IF #Stored = 0 THEN RETURN; END_IF;
    "FRK_PersistImages".D006.Rows[11] := "FRK_ConfigStore".Rows[#Stored];
    #Stored := "FRK_ConfigFind"(Scope := 'StationB.Satellite.Cell', Key := 'preset', ModelCode := 'MODEL_A');
    IF #Stored = 0 THEN RETURN; END_IF;
    "FRK_PersistImages".D006.Rows[12] := "FRK_ConfigStore".Rows[#Stored];
    #Stored := "FRK_ConfigFind"(Scope := 'StationB.Satellite.Cell.Clamp', Key := 'timeout', ModelCode := 'MODEL_A');
    IF #Stored = 0 THEN RETURN; END_IF;
    "FRK_PersistImages".D006.Rows[13] := "FRK_ConfigStore".Rows[#Stored];
    #Stored := "FRK_ConfigFind"(Scope := 'StationB.Satellite.Cell.Clamp', Key := 'preset', ModelCode := 'MODEL_A');
    IF #Stored = 0 THEN RETURN; END_IF;
    "FRK_PersistImages".D006.Rows[14] := "FRK_ConfigStore".Rows[#Stored];
    #Stored := "FRK_ConfigFind"(Scope := 'StationB.Satellite.Cell.Gate', Key := 'timeout', ModelCode := 'MODEL_A');
    IF #Stored = 0 THEN RETURN; END_IF;
    "FRK_PersistImages".D006.Rows[15] := "FRK_ConfigStore".Rows[#Stored];
    #Stored := "FRK_ConfigFind"(Scope := 'StationB.Satellite.Cell.Gate', Key := 'preset', ModelCode := 'MODEL_A');
    IF #Stored = 0 THEN RETURN; END_IF;
    "FRK_PersistImages".D006.Rows[16] := "FRK_ConfigStore".Rows[#Stored];
    #Stored := "FRK_ConfigFind"(Scope := 'StationB.Satellite.Inner', Key := 'timeout', ModelCode := 'MODEL_A');
    IF #Stored = 0 THEN RETURN; END_IF;
    "FRK_PersistImages".D006.Rows[17] := "FRK_ConfigStore".Rows[#Stored];
    #Stored := "FRK_ConfigFind"(Scope := 'StationB.Satellite.Inner', Key := 'preset', ModelCode := 'MODEL_A');
    IF #Stored = 0 THEN RETURN; END_IF;
    "FRK_PersistImages".D006.Rows[18] := "FRK_ConfigStore".Rows[#Stored];
    #Stored := "FRK_ConfigFind"(Scope := 'StationB.Satellite.Inner.Cell', Key := 'timeout', ModelCode := 'MODEL_A');
    IF #Stored = 0 THEN RETURN; END_IF;
    "FRK_PersistImages".D006.Rows[19] := "FRK_ConfigStore".Rows[#Stored];
    #Stored := "FRK_ConfigFind"(Scope := 'StationB.Satellite.Inner.Cell', Key := 'preset', ModelCode := 'MODEL_A');
    IF #Stored = 0 THEN RETURN; END_IF;
    "FRK_PersistImages".D006.Rows[20] := "FRK_ConfigStore".Rows[#Stored];
    #Stored := "FRK_ConfigFind"(Scope := 'StationB.Satellite.Inner.Cell.Clamp', Key := 'timeout', ModelCode := 'MODEL_A');
    IF #Stored = 0 THEN RETURN; END_IF;
    "FRK_PersistImages".D006.Rows[21] := "FRK_ConfigStore".Rows[#Stored];
    #Stored := "FRK_ConfigFind"(Scope := 'StationB.Satellite.Inner.Cell.Clamp', Key := 'preset', ModelCode := 'MODEL_A');
    IF #Stored = 0 THEN RETURN; END_IF;
    "FRK_PersistImages".D006.Rows[22] := "FRK_ConfigStore".Rows[#Stored];
    #Stored := "FRK_ConfigFind"(Scope := 'StationB.Satellite.Inner.Cell.Gate', Key := 'timeout', ModelCode := 'MODEL_A');
    IF #Stored = 0 THEN RETURN; END_IF;
    "FRK_PersistImages".D006.Rows[23] := "FRK_ConfigStore".Rows[#Stored];
    #Stored := "FRK_ConfigFind"(Scope := 'StationB.Satellite.Inner.Cell.Gate', Key := 'preset', ModelCode := 'MODEL_A');
    IF #Stored = 0 THEN RETURN; END_IF;
    "FRK_PersistImages".D006.Rows[24] := "FRK_ConfigStore".Rows[#Stored];
    FOR #Index := 0 TO 11401 DO "FRK_PersistBuffers".D006Data[#Index] := BYTE#0; END_FOR;
    #Position := 24;
    #NativeResult := Serialize(SRC_VARIABLE := "FRK_PersistImages".D006, DEST_ARRAY => "FRK_PersistBuffers".D006Data, POS := #Position);
    IF #NativeResult <> 0 OR #Position < 24 OR #Position > 11402 THEN RETURN; END_IF;
    #Length := #Position - 24;
    #FRK_DocCapture_D006 := TRUE;
END_FUNCTION
FUNCTION "FRK_DocApply_D006" : Bool
{ S7_Optimized_Access := 'TRUE' }
VERSION : 0.1
VAR_TEMP
    Index : Int;
    Stored : Int;
    Position : DInt;
    NativeResult : Int;
    Ok : Bool;
END_VAR
BEGIN
    #FRK_DocApply_D006 := FALSE;
    #Position := 24;
    #NativeResult := Deserialize(SRC_ARRAY := "FRK_PersistBuffers".D006Data, DEST_VARIABLE => "FRK_PersistImages".D006, POS := #Position);
    IF #NativeResult <> 0 OR #Position <> 24 + UDINT_TO_DINT("FRK_PersistConsumers".Rows[6].Result.Length) THEN RETURN; END_IF;
    IF "FRK_PersistImages".D006.SchemaVersion <> 1 OR "FRK_PersistImages".D006.Scope <> 'StationB' THEN RETURN; END_IF;
    IF "FRK_PersistImages".D006.Kind <> 0 OR "FRK_PersistImages".D006.ModelCode <> 'MODEL_A' OR "FRK_PersistImages".D006.Count <> 24 THEN RETURN; END_IF;
    IF "FRK_PersistImages".D006.ActiveModel <> 'MODEL_A' AND "FRK_PersistImages".D006.ActiveModel <> 'MODEL_B' THEN RETURN; END_IF;
    IF NOT "FRK_PersistImages".D006.Rows[1].Used OR "FRK_PersistImages".D006.Rows[1].SchemaVersion <> 4 OR "FRK_PersistImages".D006.Rows[1].ModelCode <> 'MODEL_A' OR "FRK_PersistImages".D006.Rows[1].Record.Scope <> 'StationB' OR "FRK_PersistImages".D006.Rows[1].Record.WriteKey <> 'timeout' OR "FRK_PersistImages".D006.Rows[1].Record.Revision <> 1 OR "FRK_PersistImages".D006.Rows[1].Record.Kind <> 0 OR "FRK_PersistImages".D006.Rows[1].Record.ValueType <> 3 THEN RETURN; END_IF;
    #Ok := "FRK_ConfigDecode"(Text := STRING_TO_WSTRING("FRK_PersistImages".D006.Rows[1].Record.ValueText), Storage := 7, Minimum := 1.0, Maximum := 60000.0, MaxLength := 0, Value := "FRK_ConfigScratch".Value);
    IF NOT #Ok THEN RETURN; END_IF;
    IF NOT "FRK_PersistImages".D006.Rows[2].Used OR "FRK_PersistImages".D006.Rows[2].SchemaVersion <> 4 OR "FRK_PersistImages".D006.Rows[2].ModelCode <> 'MODEL_A' OR "FRK_PersistImages".D006.Rows[2].Record.Scope <> 'StationB' OR "FRK_PersistImages".D006.Rows[2].Record.WriteKey <> 'preset' OR "FRK_PersistImages".D006.Rows[2].Record.Revision <> 2 OR "FRK_PersistImages".D006.Rows[2].Record.Kind <> 0 OR "FRK_PersistImages".D006.Rows[2].Record.ValueType <> 0 THEN RETURN; END_IF;
    #Ok := "FRK_ConfigDecode"(Text := STRING_TO_WSTRING("FRK_PersistImages".D006.Rows[2].Record.ValueText), Storage := 3, Minimum := 0.0, Maximum := 1000.0, MaxLength := 0, Value := "FRK_ConfigScratch".Value);
    IF NOT #Ok THEN RETURN; END_IF;
    IF NOT "FRK_PersistImages".D006.Rows[3].Used OR "FRK_PersistImages".D006.Rows[3].SchemaVersion <> 4 OR "FRK_PersistImages".D006.Rows[3].ModelCode <> 'MODEL_A' OR "FRK_PersistImages".D006.Rows[3].Record.Scope <> 'StationB.Cell' OR "FRK_PersistImages".D006.Rows[3].Record.WriteKey <> 'timeout' OR "FRK_PersistImages".D006.Rows[3].Record.Revision <> 1 OR "FRK_PersistImages".D006.Rows[3].Record.Kind <> 0 OR "FRK_PersistImages".D006.Rows[3].Record.ValueType <> 3 THEN RETURN; END_IF;
    #Ok := "FRK_ConfigDecode"(Text := STRING_TO_WSTRING("FRK_PersistImages".D006.Rows[3].Record.ValueText), Storage := 7, Minimum := 1.0, Maximum := 60000.0, MaxLength := 0, Value := "FRK_ConfigScratch".Value);
    IF NOT #Ok THEN RETURN; END_IF;
    IF NOT "FRK_PersistImages".D006.Rows[4].Used OR "FRK_PersistImages".D006.Rows[4].SchemaVersion <> 4 OR "FRK_PersistImages".D006.Rows[4].ModelCode <> 'MODEL_A' OR "FRK_PersistImages".D006.Rows[4].Record.Scope <> 'StationB.Cell' OR "FRK_PersistImages".D006.Rows[4].Record.WriteKey <> 'preset' OR "FRK_PersistImages".D006.Rows[4].Record.Revision <> 2 OR "FRK_PersistImages".D006.Rows[4].Record.Kind <> 0 OR "FRK_PersistImages".D006.Rows[4].Record.ValueType <> 0 THEN RETURN; END_IF;
    #Ok := "FRK_ConfigDecode"(Text := STRING_TO_WSTRING("FRK_PersistImages".D006.Rows[4].Record.ValueText), Storage := 3, Minimum := 0.0, Maximum := 1000.0, MaxLength := 0, Value := "FRK_ConfigScratch".Value);
    IF NOT #Ok THEN RETURN; END_IF;
    IF NOT "FRK_PersistImages".D006.Rows[5].Used OR "FRK_PersistImages".D006.Rows[5].SchemaVersion <> 4 OR "FRK_PersistImages".D006.Rows[5].ModelCode <> 'MODEL_A' OR "FRK_PersistImages".D006.Rows[5].Record.Scope <> 'StationB.Cell.Clamp' OR "FRK_PersistImages".D006.Rows[5].Record.WriteKey <> 'timeout' OR "FRK_PersistImages".D006.Rows[5].Record.Revision <> 1 OR "FRK_PersistImages".D006.Rows[5].Record.Kind <> 0 OR "FRK_PersistImages".D006.Rows[5].Record.ValueType <> 3 THEN RETURN; END_IF;
    #Ok := "FRK_ConfigDecode"(Text := STRING_TO_WSTRING("FRK_PersistImages".D006.Rows[5].Record.ValueText), Storage := 7, Minimum := 1.0, Maximum := 60000.0, MaxLength := 0, Value := "FRK_ConfigScratch".Value);
    IF NOT #Ok THEN RETURN; END_IF;
    IF NOT "FRK_PersistImages".D006.Rows[6].Used OR "FRK_PersistImages".D006.Rows[6].SchemaVersion <> 4 OR "FRK_PersistImages".D006.Rows[6].ModelCode <> 'MODEL_A' OR "FRK_PersistImages".D006.Rows[6].Record.Scope <> 'StationB.Cell.Clamp' OR "FRK_PersistImages".D006.Rows[6].Record.WriteKey <> 'preset' OR "FRK_PersistImages".D006.Rows[6].Record.Revision <> 2 OR "FRK_PersistImages".D006.Rows[6].Record.Kind <> 0 OR "FRK_PersistImages".D006.Rows[6].Record.ValueType <> 0 THEN RETURN; END_IF;
    #Ok := "FRK_ConfigDecode"(Text := STRING_TO_WSTRING("FRK_PersistImages".D006.Rows[6].Record.ValueText), Storage := 3, Minimum := 0.0, Maximum := 1000.0, MaxLength := 0, Value := "FRK_ConfigScratch".Value);
    IF NOT #Ok THEN RETURN; END_IF;
    IF NOT "FRK_PersistImages".D006.Rows[7].Used OR "FRK_PersistImages".D006.Rows[7].SchemaVersion <> 4 OR "FRK_PersistImages".D006.Rows[7].ModelCode <> 'MODEL_A' OR "FRK_PersistImages".D006.Rows[7].Record.Scope <> 'StationB.Cell.Gate' OR "FRK_PersistImages".D006.Rows[7].Record.WriteKey <> 'timeout' OR "FRK_PersistImages".D006.Rows[7].Record.Revision <> 1 OR "FRK_PersistImages".D006.Rows[7].Record.Kind <> 0 OR "FRK_PersistImages".D006.Rows[7].Record.ValueType <> 3 THEN RETURN; END_IF;
    #Ok := "FRK_ConfigDecode"(Text := STRING_TO_WSTRING("FRK_PersistImages".D006.Rows[7].Record.ValueText), Storage := 7, Minimum := 1.0, Maximum := 60000.0, MaxLength := 0, Value := "FRK_ConfigScratch".Value);
    IF NOT #Ok THEN RETURN; END_IF;
    IF NOT "FRK_PersistImages".D006.Rows[8].Used OR "FRK_PersistImages".D006.Rows[8].SchemaVersion <> 4 OR "FRK_PersistImages".D006.Rows[8].ModelCode <> 'MODEL_A' OR "FRK_PersistImages".D006.Rows[8].Record.Scope <> 'StationB.Cell.Gate' OR "FRK_PersistImages".D006.Rows[8].Record.WriteKey <> 'preset' OR "FRK_PersistImages".D006.Rows[8].Record.Revision <> 2 OR "FRK_PersistImages".D006.Rows[8].Record.Kind <> 0 OR "FRK_PersistImages".D006.Rows[8].Record.ValueType <> 0 THEN RETURN; END_IF;
    #Ok := "FRK_ConfigDecode"(Text := STRING_TO_WSTRING("FRK_PersistImages".D006.Rows[8].Record.ValueText), Storage := 3, Minimum := 0.0, Maximum := 1000.0, MaxLength := 0, Value := "FRK_ConfigScratch".Value);
    IF NOT #Ok THEN RETURN; END_IF;
    IF NOT "FRK_PersistImages".D006.Rows[9].Used OR "FRK_PersistImages".D006.Rows[9].SchemaVersion <> 4 OR "FRK_PersistImages".D006.Rows[9].ModelCode <> 'MODEL_A' OR "FRK_PersistImages".D006.Rows[9].Record.Scope <> 'StationB.Satellite' OR "FRK_PersistImages".D006.Rows[9].Record.WriteKey <> 'timeout' OR "FRK_PersistImages".D006.Rows[9].Record.Revision <> 1 OR "FRK_PersistImages".D006.Rows[9].Record.Kind <> 0 OR "FRK_PersistImages".D006.Rows[9].Record.ValueType <> 3 THEN RETURN; END_IF;
    #Ok := "FRK_ConfigDecode"(Text := STRING_TO_WSTRING("FRK_PersistImages".D006.Rows[9].Record.ValueText), Storage := 7, Minimum := 1.0, Maximum := 60000.0, MaxLength := 0, Value := "FRK_ConfigScratch".Value);
    IF NOT #Ok THEN RETURN; END_IF;
    IF NOT "FRK_PersistImages".D006.Rows[10].Used OR "FRK_PersistImages".D006.Rows[10].SchemaVersion <> 4 OR "FRK_PersistImages".D006.Rows[10].ModelCode <> 'MODEL_A' OR "FRK_PersistImages".D006.Rows[10].Record.Scope <> 'StationB.Satellite' OR "FRK_PersistImages".D006.Rows[10].Record.WriteKey <> 'preset' OR "FRK_PersistImages".D006.Rows[10].Record.Revision <> 2 OR "FRK_PersistImages".D006.Rows[10].Record.Kind <> 0 OR "FRK_PersistImages".D006.Rows[10].Record.ValueType <> 0 THEN RETURN; END_IF;
    #Ok := "FRK_ConfigDecode"(Text := STRING_TO_WSTRING("FRK_PersistImages".D006.Rows[10].Record.ValueText), Storage := 3, Minimum := 0.0, Maximum := 1000.0, MaxLength := 0, Value := "FRK_ConfigScratch".Value);
    IF NOT #Ok THEN RETURN; END_IF;
    IF NOT "FRK_PersistImages".D006.Rows[11].Used OR "FRK_PersistImages".D006.Rows[11].SchemaVersion <> 4 OR "FRK_PersistImages".D006.Rows[11].ModelCode <> 'MODEL_A' OR "FRK_PersistImages".D006.Rows[11].Record.Scope <> 'StationB.Satellite.Cell' OR "FRK_PersistImages".D006.Rows[11].Record.WriteKey <> 'timeout' OR "FRK_PersistImages".D006.Rows[11].Record.Revision <> 1 OR "FRK_PersistImages".D006.Rows[11].Record.Kind <> 0 OR "FRK_PersistImages".D006.Rows[11].Record.ValueType <> 3 THEN RETURN; END_IF;
    #Ok := "FRK_ConfigDecode"(Text := STRING_TO_WSTRING("FRK_PersistImages".D006.Rows[11].Record.ValueText), Storage := 7, Minimum := 1.0, Maximum := 60000.0, MaxLength := 0, Value := "FRK_ConfigScratch".Value);
    IF NOT #Ok THEN RETURN; END_IF;
    IF NOT "FRK_PersistImages".D006.Rows[12].Used OR "FRK_PersistImages".D006.Rows[12].SchemaVersion <> 4 OR "FRK_PersistImages".D006.Rows[12].ModelCode <> 'MODEL_A' OR "FRK_PersistImages".D006.Rows[12].Record.Scope <> 'StationB.Satellite.Cell' OR "FRK_PersistImages".D006.Rows[12].Record.WriteKey <> 'preset' OR "FRK_PersistImages".D006.Rows[12].Record.Revision <> 2 OR "FRK_PersistImages".D006.Rows[12].Record.Kind <> 0 OR "FRK_PersistImages".D006.Rows[12].Record.ValueType <> 0 THEN RETURN; END_IF;
    #Ok := "FRK_ConfigDecode"(Text := STRING_TO_WSTRING("FRK_PersistImages".D006.Rows[12].Record.ValueText), Storage := 3, Minimum := 0.0, Maximum := 1000.0, MaxLength := 0, Value := "FRK_ConfigScratch".Value);
    IF NOT #Ok THEN RETURN; END_IF;
    IF NOT "FRK_PersistImages".D006.Rows[13].Used OR "FRK_PersistImages".D006.Rows[13].SchemaVersion <> 4 OR "FRK_PersistImages".D006.Rows[13].ModelCode <> 'MODEL_A' OR "FRK_PersistImages".D006.Rows[13].Record.Scope <> 'StationB.Satellite.Cell.Clamp' OR "FRK_PersistImages".D006.Rows[13].Record.WriteKey <> 'timeout' OR "FRK_PersistImages".D006.Rows[13].Record.Revision <> 1 OR "FRK_PersistImages".D006.Rows[13].Record.Kind <> 0 OR "FRK_PersistImages".D006.Rows[13].Record.ValueType <> 3 THEN RETURN; END_IF;
    #Ok := "FRK_ConfigDecode"(Text := STRING_TO_WSTRING("FRK_PersistImages".D006.Rows[13].Record.ValueText), Storage := 7, Minimum := 1.0, Maximum := 60000.0, MaxLength := 0, Value := "FRK_ConfigScratch".Value);
    IF NOT #Ok THEN RETURN; END_IF;
    IF NOT "FRK_PersistImages".D006.Rows[14].Used OR "FRK_PersistImages".D006.Rows[14].SchemaVersion <> 4 OR "FRK_PersistImages".D006.Rows[14].ModelCode <> 'MODEL_A' OR "FRK_PersistImages".D006.Rows[14].Record.Scope <> 'StationB.Satellite.Cell.Clamp' OR "FRK_PersistImages".D006.Rows[14].Record.WriteKey <> 'preset' OR "FRK_PersistImages".D006.Rows[14].Record.Revision <> 2 OR "FRK_PersistImages".D006.Rows[14].Record.Kind <> 0 OR "FRK_PersistImages".D006.Rows[14].Record.ValueType <> 0 THEN RETURN; END_IF;
    #Ok := "FRK_ConfigDecode"(Text := STRING_TO_WSTRING("FRK_PersistImages".D006.Rows[14].Record.ValueText), Storage := 3, Minimum := 0.0, Maximum := 1000.0, MaxLength := 0, Value := "FRK_ConfigScratch".Value);
    IF NOT #Ok THEN RETURN; END_IF;
    IF NOT "FRK_PersistImages".D006.Rows[15].Used OR "FRK_PersistImages".D006.Rows[15].SchemaVersion <> 4 OR "FRK_PersistImages".D006.Rows[15].ModelCode <> 'MODEL_A' OR "FRK_PersistImages".D006.Rows[15].Record.Scope <> 'StationB.Satellite.Cell.Gate' OR "FRK_PersistImages".D006.Rows[15].Record.WriteKey <> 'timeout' OR "FRK_PersistImages".D006.Rows[15].Record.Revision <> 1 OR "FRK_PersistImages".D006.Rows[15].Record.Kind <> 0 OR "FRK_PersistImages".D006.Rows[15].Record.ValueType <> 3 THEN RETURN; END_IF;
    #Ok := "FRK_ConfigDecode"(Text := STRING_TO_WSTRING("FRK_PersistImages".D006.Rows[15].Record.ValueText), Storage := 7, Minimum := 1.0, Maximum := 60000.0, MaxLength := 0, Value := "FRK_ConfigScratch".Value);
    IF NOT #Ok THEN RETURN; END_IF;
    IF NOT "FRK_PersistImages".D006.Rows[16].Used OR "FRK_PersistImages".D006.Rows[16].SchemaVersion <> 4 OR "FRK_PersistImages".D006.Rows[16].ModelCode <> 'MODEL_A' OR "FRK_PersistImages".D006.Rows[16].Record.Scope <> 'StationB.Satellite.Cell.Gate' OR "FRK_PersistImages".D006.Rows[16].Record.WriteKey <> 'preset' OR "FRK_PersistImages".D006.Rows[16].Record.Revision <> 2 OR "FRK_PersistImages".D006.Rows[16].Record.Kind <> 0 OR "FRK_PersistImages".D006.Rows[16].Record.ValueType <> 0 THEN RETURN; END_IF;
    #Ok := "FRK_ConfigDecode"(Text := STRING_TO_WSTRING("FRK_PersistImages".D006.Rows[16].Record.ValueText), Storage := 3, Minimum := 0.0, Maximum := 1000.0, MaxLength := 0, Value := "FRK_ConfigScratch".Value);
    IF NOT #Ok THEN RETURN; END_IF;
    IF NOT "FRK_PersistImages".D006.Rows[17].Used OR "FRK_PersistImages".D006.Rows[17].SchemaVersion <> 4 OR "FRK_PersistImages".D006.Rows[17].ModelCode <> 'MODEL_A' OR "FRK_PersistImages".D006.Rows[17].Record.Scope <> 'StationB.Satellite.Inner' OR "FRK_PersistImages".D006.Rows[17].Record.WriteKey <> 'timeout' OR "FRK_PersistImages".D006.Rows[17].Record.Revision <> 1 OR "FRK_PersistImages".D006.Rows[17].Record.Kind <> 0 OR "FRK_PersistImages".D006.Rows[17].Record.ValueType <> 3 THEN RETURN; END_IF;
    #Ok := "FRK_ConfigDecode"(Text := STRING_TO_WSTRING("FRK_PersistImages".D006.Rows[17].Record.ValueText), Storage := 7, Minimum := 1.0, Maximum := 60000.0, MaxLength := 0, Value := "FRK_ConfigScratch".Value);
    IF NOT #Ok THEN RETURN; END_IF;
    IF NOT "FRK_PersistImages".D006.Rows[18].Used OR "FRK_PersistImages".D006.Rows[18].SchemaVersion <> 4 OR "FRK_PersistImages".D006.Rows[18].ModelCode <> 'MODEL_A' OR "FRK_PersistImages".D006.Rows[18].Record.Scope <> 'StationB.Satellite.Inner' OR "FRK_PersistImages".D006.Rows[18].Record.WriteKey <> 'preset' OR "FRK_PersistImages".D006.Rows[18].Record.Revision <> 2 OR "FRK_PersistImages".D006.Rows[18].Record.Kind <> 0 OR "FRK_PersistImages".D006.Rows[18].Record.ValueType <> 0 THEN RETURN; END_IF;
    #Ok := "FRK_ConfigDecode"(Text := STRING_TO_WSTRING("FRK_PersistImages".D006.Rows[18].Record.ValueText), Storage := 3, Minimum := 0.0, Maximum := 1000.0, MaxLength := 0, Value := "FRK_ConfigScratch".Value);
    IF NOT #Ok THEN RETURN; END_IF;
    IF NOT "FRK_PersistImages".D006.Rows[19].Used OR "FRK_PersistImages".D006.Rows[19].SchemaVersion <> 4 OR "FRK_PersistImages".D006.Rows[19].ModelCode <> 'MODEL_A' OR "FRK_PersistImages".D006.Rows[19].Record.Scope <> 'StationB.Satellite.Inner.Cell' OR "FRK_PersistImages".D006.Rows[19].Record.WriteKey <> 'timeout' OR "FRK_PersistImages".D006.Rows[19].Record.Revision <> 1 OR "FRK_PersistImages".D006.Rows[19].Record.Kind <> 0 OR "FRK_PersistImages".D006.Rows[19].Record.ValueType <> 3 THEN RETURN; END_IF;
    #Ok := "FRK_ConfigDecode"(Text := STRING_TO_WSTRING("FRK_PersistImages".D006.Rows[19].Record.ValueText), Storage := 7, Minimum := 1.0, Maximum := 60000.0, MaxLength := 0, Value := "FRK_ConfigScratch".Value);
    IF NOT #Ok THEN RETURN; END_IF;
    IF NOT "FRK_PersistImages".D006.Rows[20].Used OR "FRK_PersistImages".D006.Rows[20].SchemaVersion <> 4 OR "FRK_PersistImages".D006.Rows[20].ModelCode <> 'MODEL_A' OR "FRK_PersistImages".D006.Rows[20].Record.Scope <> 'StationB.Satellite.Inner.Cell' OR "FRK_PersistImages".D006.Rows[20].Record.WriteKey <> 'preset' OR "FRK_PersistImages".D006.Rows[20].Record.Revision <> 2 OR "FRK_PersistImages".D006.Rows[20].Record.Kind <> 0 OR "FRK_PersistImages".D006.Rows[20].Record.ValueType <> 0 THEN RETURN; END_IF;
    #Ok := "FRK_ConfigDecode"(Text := STRING_TO_WSTRING("FRK_PersistImages".D006.Rows[20].Record.ValueText), Storage := 3, Minimum := 0.0, Maximum := 1000.0, MaxLength := 0, Value := "FRK_ConfigScratch".Value);
    IF NOT #Ok THEN RETURN; END_IF;
    IF NOT "FRK_PersistImages".D006.Rows[21].Used OR "FRK_PersistImages".D006.Rows[21].SchemaVersion <> 4 OR "FRK_PersistImages".D006.Rows[21].ModelCode <> 'MODEL_A' OR "FRK_PersistImages".D006.Rows[21].Record.Scope <> 'StationB.Satellite.Inner.Cell.Clamp' OR "FRK_PersistImages".D006.Rows[21].Record.WriteKey <> 'timeout' OR "FRK_PersistImages".D006.Rows[21].Record.Revision <> 1 OR "FRK_PersistImages".D006.Rows[21].Record.Kind <> 0 OR "FRK_PersistImages".D006.Rows[21].Record.ValueType <> 3 THEN RETURN; END_IF;
    #Ok := "FRK_ConfigDecode"(Text := STRING_TO_WSTRING("FRK_PersistImages".D006.Rows[21].Record.ValueText), Storage := 7, Minimum := 1.0, Maximum := 60000.0, MaxLength := 0, Value := "FRK_ConfigScratch".Value);
    IF NOT #Ok THEN RETURN; END_IF;
    IF NOT "FRK_PersistImages".D006.Rows[22].Used OR "FRK_PersistImages".D006.Rows[22].SchemaVersion <> 4 OR "FRK_PersistImages".D006.Rows[22].ModelCode <> 'MODEL_A' OR "FRK_PersistImages".D006.Rows[22].Record.Scope <> 'StationB.Satellite.Inner.Cell.Clamp' OR "FRK_PersistImages".D006.Rows[22].Record.WriteKey <> 'preset' OR "FRK_PersistImages".D006.Rows[22].Record.Revision <> 2 OR "FRK_PersistImages".D006.Rows[22].Record.Kind <> 0 OR "FRK_PersistImages".D006.Rows[22].Record.ValueType <> 0 THEN RETURN; END_IF;
    #Ok := "FRK_ConfigDecode"(Text := STRING_TO_WSTRING("FRK_PersistImages".D006.Rows[22].Record.ValueText), Storage := 3, Minimum := 0.0, Maximum := 1000.0, MaxLength := 0, Value := "FRK_ConfigScratch".Value);
    IF NOT #Ok THEN RETURN; END_IF;
    IF NOT "FRK_PersistImages".D006.Rows[23].Used OR "FRK_PersistImages".D006.Rows[23].SchemaVersion <> 4 OR "FRK_PersistImages".D006.Rows[23].ModelCode <> 'MODEL_A' OR "FRK_PersistImages".D006.Rows[23].Record.Scope <> 'StationB.Satellite.Inner.Cell.Gate' OR "FRK_PersistImages".D006.Rows[23].Record.WriteKey <> 'timeout' OR "FRK_PersistImages".D006.Rows[23].Record.Revision <> 1 OR "FRK_PersistImages".D006.Rows[23].Record.Kind <> 0 OR "FRK_PersistImages".D006.Rows[23].Record.ValueType <> 3 THEN RETURN; END_IF;
    #Ok := "FRK_ConfigDecode"(Text := STRING_TO_WSTRING("FRK_PersistImages".D006.Rows[23].Record.ValueText), Storage := 7, Minimum := 1.0, Maximum := 60000.0, MaxLength := 0, Value := "FRK_ConfigScratch".Value);
    IF NOT #Ok THEN RETURN; END_IF;
    IF NOT "FRK_PersistImages".D006.Rows[24].Used OR "FRK_PersistImages".D006.Rows[24].SchemaVersion <> 4 OR "FRK_PersistImages".D006.Rows[24].ModelCode <> 'MODEL_A' OR "FRK_PersistImages".D006.Rows[24].Record.Scope <> 'StationB.Satellite.Inner.Cell.Gate' OR "FRK_PersistImages".D006.Rows[24].Record.WriteKey <> 'preset' OR "FRK_PersistImages".D006.Rows[24].Record.Revision <> 2 OR "FRK_PersistImages".D006.Rows[24].Record.Kind <> 0 OR "FRK_PersistImages".D006.Rows[24].Record.ValueType <> 0 THEN RETURN; END_IF;
    #Ok := "FRK_ConfigDecode"(Text := STRING_TO_WSTRING("FRK_PersistImages".D006.Rows[24].Record.ValueText), Storage := 3, Minimum := 0.0, Maximum := 1000.0, MaxLength := 0, Value := "FRK_ConfigScratch".Value);
    IF NOT #Ok THEN RETURN; END_IF;
    #Stored := "FRK_ConfigFind"(Scope := 'StationB', Key := 'timeout', ModelCode := 'MODEL_A');
    IF #Stored = 0 THEN
        FOR #Stored := 1 TO 108 DO IF NOT "FRK_ConfigStore".Rows[#Stored].Used THEN EXIT; END_IF; END_FOR;
    END_IF;
    IF #Stored < 1 OR #Stored > 108 THEN RETURN; END_IF;
    "FRK_ConfigStore".Rows[#Stored] := "FRK_PersistImages".D006.Rows[1];
    #Stored := "FRK_ConfigFind"(Scope := 'StationB', Key := 'preset', ModelCode := 'MODEL_A');
    IF #Stored = 0 THEN
        FOR #Stored := 1 TO 108 DO IF NOT "FRK_ConfigStore".Rows[#Stored].Used THEN EXIT; END_IF; END_FOR;
    END_IF;
    IF #Stored < 1 OR #Stored > 108 THEN RETURN; END_IF;
    "FRK_ConfigStore".Rows[#Stored] := "FRK_PersistImages".D006.Rows[2];
    #Stored := "FRK_ConfigFind"(Scope := 'StationB.Cell', Key := 'timeout', ModelCode := 'MODEL_A');
    IF #Stored = 0 THEN
        FOR #Stored := 1 TO 108 DO IF NOT "FRK_ConfigStore".Rows[#Stored].Used THEN EXIT; END_IF; END_FOR;
    END_IF;
    IF #Stored < 1 OR #Stored > 108 THEN RETURN; END_IF;
    "FRK_ConfigStore".Rows[#Stored] := "FRK_PersistImages".D006.Rows[3];
    #Stored := "FRK_ConfigFind"(Scope := 'StationB.Cell', Key := 'preset', ModelCode := 'MODEL_A');
    IF #Stored = 0 THEN
        FOR #Stored := 1 TO 108 DO IF NOT "FRK_ConfigStore".Rows[#Stored].Used THEN EXIT; END_IF; END_FOR;
    END_IF;
    IF #Stored < 1 OR #Stored > 108 THEN RETURN; END_IF;
    "FRK_ConfigStore".Rows[#Stored] := "FRK_PersistImages".D006.Rows[4];
    #Stored := "FRK_ConfigFind"(Scope := 'StationB.Cell.Clamp', Key := 'timeout', ModelCode := 'MODEL_A');
    IF #Stored = 0 THEN
        FOR #Stored := 1 TO 108 DO IF NOT "FRK_ConfigStore".Rows[#Stored].Used THEN EXIT; END_IF; END_FOR;
    END_IF;
    IF #Stored < 1 OR #Stored > 108 THEN RETURN; END_IF;
    "FRK_ConfigStore".Rows[#Stored] := "FRK_PersistImages".D006.Rows[5];
    #Stored := "FRK_ConfigFind"(Scope := 'StationB.Cell.Clamp', Key := 'preset', ModelCode := 'MODEL_A');
    IF #Stored = 0 THEN
        FOR #Stored := 1 TO 108 DO IF NOT "FRK_ConfigStore".Rows[#Stored].Used THEN EXIT; END_IF; END_FOR;
    END_IF;
    IF #Stored < 1 OR #Stored > 108 THEN RETURN; END_IF;
    "FRK_ConfigStore".Rows[#Stored] := "FRK_PersistImages".D006.Rows[6];
    #Stored := "FRK_ConfigFind"(Scope := 'StationB.Cell.Gate', Key := 'timeout', ModelCode := 'MODEL_A');
    IF #Stored = 0 THEN
        FOR #Stored := 1 TO 108 DO IF NOT "FRK_ConfigStore".Rows[#Stored].Used THEN EXIT; END_IF; END_FOR;
    END_IF;
    IF #Stored < 1 OR #Stored > 108 THEN RETURN; END_IF;
    "FRK_ConfigStore".Rows[#Stored] := "FRK_PersistImages".D006.Rows[7];
    #Stored := "FRK_ConfigFind"(Scope := 'StationB.Cell.Gate', Key := 'preset', ModelCode := 'MODEL_A');
    IF #Stored = 0 THEN
        FOR #Stored := 1 TO 108 DO IF NOT "FRK_ConfigStore".Rows[#Stored].Used THEN EXIT; END_IF; END_FOR;
    END_IF;
    IF #Stored < 1 OR #Stored > 108 THEN RETURN; END_IF;
    "FRK_ConfigStore".Rows[#Stored] := "FRK_PersistImages".D006.Rows[8];
    #Stored := "FRK_ConfigFind"(Scope := 'StationB.Satellite', Key := 'timeout', ModelCode := 'MODEL_A');
    IF #Stored = 0 THEN
        FOR #Stored := 1 TO 108 DO IF NOT "FRK_ConfigStore".Rows[#Stored].Used THEN EXIT; END_IF; END_FOR;
    END_IF;
    IF #Stored < 1 OR #Stored > 108 THEN RETURN; END_IF;
    "FRK_ConfigStore".Rows[#Stored] := "FRK_PersistImages".D006.Rows[9];
    #Stored := "FRK_ConfigFind"(Scope := 'StationB.Satellite', Key := 'preset', ModelCode := 'MODEL_A');
    IF #Stored = 0 THEN
        FOR #Stored := 1 TO 108 DO IF NOT "FRK_ConfigStore".Rows[#Stored].Used THEN EXIT; END_IF; END_FOR;
    END_IF;
    IF #Stored < 1 OR #Stored > 108 THEN RETURN; END_IF;
    "FRK_ConfigStore".Rows[#Stored] := "FRK_PersistImages".D006.Rows[10];
    #Stored := "FRK_ConfigFind"(Scope := 'StationB.Satellite.Cell', Key := 'timeout', ModelCode := 'MODEL_A');
    IF #Stored = 0 THEN
        FOR #Stored := 1 TO 108 DO IF NOT "FRK_ConfigStore".Rows[#Stored].Used THEN EXIT; END_IF; END_FOR;
    END_IF;
    IF #Stored < 1 OR #Stored > 108 THEN RETURN; END_IF;
    "FRK_ConfigStore".Rows[#Stored] := "FRK_PersistImages".D006.Rows[11];
    #Stored := "FRK_ConfigFind"(Scope := 'StationB.Satellite.Cell', Key := 'preset', ModelCode := 'MODEL_A');
    IF #Stored = 0 THEN
        FOR #Stored := 1 TO 108 DO IF NOT "FRK_ConfigStore".Rows[#Stored].Used THEN EXIT; END_IF; END_FOR;
    END_IF;
    IF #Stored < 1 OR #Stored > 108 THEN RETURN; END_IF;
    "FRK_ConfigStore".Rows[#Stored] := "FRK_PersistImages".D006.Rows[12];
    #Stored := "FRK_ConfigFind"(Scope := 'StationB.Satellite.Cell.Clamp', Key := 'timeout', ModelCode := 'MODEL_A');
    IF #Stored = 0 THEN
        FOR #Stored := 1 TO 108 DO IF NOT "FRK_ConfigStore".Rows[#Stored].Used THEN EXIT; END_IF; END_FOR;
    END_IF;
    IF #Stored < 1 OR #Stored > 108 THEN RETURN; END_IF;
    "FRK_ConfigStore".Rows[#Stored] := "FRK_PersistImages".D006.Rows[13];
    #Stored := "FRK_ConfigFind"(Scope := 'StationB.Satellite.Cell.Clamp', Key := 'preset', ModelCode := 'MODEL_A');
    IF #Stored = 0 THEN
        FOR #Stored := 1 TO 108 DO IF NOT "FRK_ConfigStore".Rows[#Stored].Used THEN EXIT; END_IF; END_FOR;
    END_IF;
    IF #Stored < 1 OR #Stored > 108 THEN RETURN; END_IF;
    "FRK_ConfigStore".Rows[#Stored] := "FRK_PersistImages".D006.Rows[14];
    #Stored := "FRK_ConfigFind"(Scope := 'StationB.Satellite.Cell.Gate', Key := 'timeout', ModelCode := 'MODEL_A');
    IF #Stored = 0 THEN
        FOR #Stored := 1 TO 108 DO IF NOT "FRK_ConfigStore".Rows[#Stored].Used THEN EXIT; END_IF; END_FOR;
    END_IF;
    IF #Stored < 1 OR #Stored > 108 THEN RETURN; END_IF;
    "FRK_ConfigStore".Rows[#Stored] := "FRK_PersistImages".D006.Rows[15];
    #Stored := "FRK_ConfigFind"(Scope := 'StationB.Satellite.Cell.Gate', Key := 'preset', ModelCode := 'MODEL_A');
    IF #Stored = 0 THEN
        FOR #Stored := 1 TO 108 DO IF NOT "FRK_ConfigStore".Rows[#Stored].Used THEN EXIT; END_IF; END_FOR;
    END_IF;
    IF #Stored < 1 OR #Stored > 108 THEN RETURN; END_IF;
    "FRK_ConfigStore".Rows[#Stored] := "FRK_PersistImages".D006.Rows[16];
    #Stored := "FRK_ConfigFind"(Scope := 'StationB.Satellite.Inner', Key := 'timeout', ModelCode := 'MODEL_A');
    IF #Stored = 0 THEN
        FOR #Stored := 1 TO 108 DO IF NOT "FRK_ConfigStore".Rows[#Stored].Used THEN EXIT; END_IF; END_FOR;
    END_IF;
    IF #Stored < 1 OR #Stored > 108 THEN RETURN; END_IF;
    "FRK_ConfigStore".Rows[#Stored] := "FRK_PersistImages".D006.Rows[17];
    #Stored := "FRK_ConfigFind"(Scope := 'StationB.Satellite.Inner', Key := 'preset', ModelCode := 'MODEL_A');
    IF #Stored = 0 THEN
        FOR #Stored := 1 TO 108 DO IF NOT "FRK_ConfigStore".Rows[#Stored].Used THEN EXIT; END_IF; END_FOR;
    END_IF;
    IF #Stored < 1 OR #Stored > 108 THEN RETURN; END_IF;
    "FRK_ConfigStore".Rows[#Stored] := "FRK_PersistImages".D006.Rows[18];
    #Stored := "FRK_ConfigFind"(Scope := 'StationB.Satellite.Inner.Cell', Key := 'timeout', ModelCode := 'MODEL_A');
    IF #Stored = 0 THEN
        FOR #Stored := 1 TO 108 DO IF NOT "FRK_ConfigStore".Rows[#Stored].Used THEN EXIT; END_IF; END_FOR;
    END_IF;
    IF #Stored < 1 OR #Stored > 108 THEN RETURN; END_IF;
    "FRK_ConfigStore".Rows[#Stored] := "FRK_PersistImages".D006.Rows[19];
    #Stored := "FRK_ConfigFind"(Scope := 'StationB.Satellite.Inner.Cell', Key := 'preset', ModelCode := 'MODEL_A');
    IF #Stored = 0 THEN
        FOR #Stored := 1 TO 108 DO IF NOT "FRK_ConfigStore".Rows[#Stored].Used THEN EXIT; END_IF; END_FOR;
    END_IF;
    IF #Stored < 1 OR #Stored > 108 THEN RETURN; END_IF;
    "FRK_ConfigStore".Rows[#Stored] := "FRK_PersistImages".D006.Rows[20];
    #Stored := "FRK_ConfigFind"(Scope := 'StationB.Satellite.Inner.Cell.Clamp', Key := 'timeout', ModelCode := 'MODEL_A');
    IF #Stored = 0 THEN
        FOR #Stored := 1 TO 108 DO IF NOT "FRK_ConfigStore".Rows[#Stored].Used THEN EXIT; END_IF; END_FOR;
    END_IF;
    IF #Stored < 1 OR #Stored > 108 THEN RETURN; END_IF;
    "FRK_ConfigStore".Rows[#Stored] := "FRK_PersistImages".D006.Rows[21];
    #Stored := "FRK_ConfigFind"(Scope := 'StationB.Satellite.Inner.Cell.Clamp', Key := 'preset', ModelCode := 'MODEL_A');
    IF #Stored = 0 THEN
        FOR #Stored := 1 TO 108 DO IF NOT "FRK_ConfigStore".Rows[#Stored].Used THEN EXIT; END_IF; END_FOR;
    END_IF;
    IF #Stored < 1 OR #Stored > 108 THEN RETURN; END_IF;
    "FRK_ConfigStore".Rows[#Stored] := "FRK_PersistImages".D006.Rows[22];
    #Stored := "FRK_ConfigFind"(Scope := 'StationB.Satellite.Inner.Cell.Gate', Key := 'timeout', ModelCode := 'MODEL_A');
    IF #Stored = 0 THEN
        FOR #Stored := 1 TO 108 DO IF NOT "FRK_ConfigStore".Rows[#Stored].Used THEN EXIT; END_IF; END_FOR;
    END_IF;
    IF #Stored < 1 OR #Stored > 108 THEN RETURN; END_IF;
    "FRK_ConfigStore".Rows[#Stored] := "FRK_PersistImages".D006.Rows[23];
    #Stored := "FRK_ConfigFind"(Scope := 'StationB.Satellite.Inner.Cell.Gate', Key := 'preset', ModelCode := 'MODEL_A');
    IF #Stored = 0 THEN
        FOR #Stored := 1 TO 108 DO IF NOT "FRK_ConfigStore".Rows[#Stored].Used THEN EXIT; END_IF; END_FOR;
    END_IF;
    IF #Stored < 1 OR #Stored > 108 THEN RETURN; END_IF;
    "FRK_ConfigStore".Rows[#Stored] := "FRK_PersistImages".D006.Rows[24];
    "FRK_ConfigStore".SchemaVersion := 1;
    #FRK_DocApply_D006 := TRUE;
END_FUNCTION
FUNCTION "FRK_DocCapture_D007" : Bool
{ S7_Optimized_Access := 'TRUE' }
VERSION : 0.1
VAR_IN_OUT
    Length : DInt;
END_VAR
VAR_TEMP
    Index : Int;
    Stored : Int;
    Position : DInt;
    NativeResult : Int;
    Ok : Bool;
END_VAR
BEGIN
    #FRK_DocCapture_D007 := FALSE;
    "FRK_PersistImages".D007.SchemaVersion := 1; "FRK_PersistImages".D007.Scope := 'StationB';
    "FRK_PersistImages".D007.Kind := 0;
    "FRK_PersistImages".D007.ModelCode := 'MODEL_B';
    "FRK_PersistImages".D007.ActiveModel := "FRK_ConfigStore".ActiveModels[2];
    "FRK_PersistImages".D007.Count := 24;
    #Stored := "FRK_ConfigFind"(Scope := 'StationB', Key := 'timeout', ModelCode := 'MODEL_B');
    IF #Stored = 0 THEN RETURN; END_IF;
    "FRK_PersistImages".D007.Rows[1] := "FRK_ConfigStore".Rows[#Stored];
    #Stored := "FRK_ConfigFind"(Scope := 'StationB', Key := 'preset', ModelCode := 'MODEL_B');
    IF #Stored = 0 THEN RETURN; END_IF;
    "FRK_PersistImages".D007.Rows[2] := "FRK_ConfigStore".Rows[#Stored];
    #Stored := "FRK_ConfigFind"(Scope := 'StationB.Cell', Key := 'timeout', ModelCode := 'MODEL_B');
    IF #Stored = 0 THEN RETURN; END_IF;
    "FRK_PersistImages".D007.Rows[3] := "FRK_ConfigStore".Rows[#Stored];
    #Stored := "FRK_ConfigFind"(Scope := 'StationB.Cell', Key := 'preset', ModelCode := 'MODEL_B');
    IF #Stored = 0 THEN RETURN; END_IF;
    "FRK_PersistImages".D007.Rows[4] := "FRK_ConfigStore".Rows[#Stored];
    #Stored := "FRK_ConfigFind"(Scope := 'StationB.Cell.Clamp', Key := 'timeout', ModelCode := 'MODEL_B');
    IF #Stored = 0 THEN RETURN; END_IF;
    "FRK_PersistImages".D007.Rows[5] := "FRK_ConfigStore".Rows[#Stored];
    #Stored := "FRK_ConfigFind"(Scope := 'StationB.Cell.Clamp', Key := 'preset', ModelCode := 'MODEL_B');
    IF #Stored = 0 THEN RETURN; END_IF;
    "FRK_PersistImages".D007.Rows[6] := "FRK_ConfigStore".Rows[#Stored];
    #Stored := "FRK_ConfigFind"(Scope := 'StationB.Cell.Gate', Key := 'timeout', ModelCode := 'MODEL_B');
    IF #Stored = 0 THEN RETURN; END_IF;
    "FRK_PersistImages".D007.Rows[7] := "FRK_ConfigStore".Rows[#Stored];
    #Stored := "FRK_ConfigFind"(Scope := 'StationB.Cell.Gate', Key := 'preset', ModelCode := 'MODEL_B');
    IF #Stored = 0 THEN RETURN; END_IF;
    "FRK_PersistImages".D007.Rows[8] := "FRK_ConfigStore".Rows[#Stored];
    #Stored := "FRK_ConfigFind"(Scope := 'StationB.Satellite', Key := 'timeout', ModelCode := 'MODEL_B');
    IF #Stored = 0 THEN RETURN; END_IF;
    "FRK_PersistImages".D007.Rows[9] := "FRK_ConfigStore".Rows[#Stored];
    #Stored := "FRK_ConfigFind"(Scope := 'StationB.Satellite', Key := 'preset', ModelCode := 'MODEL_B');
    IF #Stored = 0 THEN RETURN; END_IF;
    "FRK_PersistImages".D007.Rows[10] := "FRK_ConfigStore".Rows[#Stored];
    #Stored := "FRK_ConfigFind"(Scope := 'StationB.Satellite.Cell', Key := 'timeout', ModelCode := 'MODEL_B');
    IF #Stored = 0 THEN RETURN; END_IF;
    "FRK_PersistImages".D007.Rows[11] := "FRK_ConfigStore".Rows[#Stored];
    #Stored := "FRK_ConfigFind"(Scope := 'StationB.Satellite.Cell', Key := 'preset', ModelCode := 'MODEL_B');
    IF #Stored = 0 THEN RETURN; END_IF;
    "FRK_PersistImages".D007.Rows[12] := "FRK_ConfigStore".Rows[#Stored];
    #Stored := "FRK_ConfigFind"(Scope := 'StationB.Satellite.Cell.Clamp', Key := 'timeout', ModelCode := 'MODEL_B');
    IF #Stored = 0 THEN RETURN; END_IF;
    "FRK_PersistImages".D007.Rows[13] := "FRK_ConfigStore".Rows[#Stored];
    #Stored := "FRK_ConfigFind"(Scope := 'StationB.Satellite.Cell.Clamp', Key := 'preset', ModelCode := 'MODEL_B');
    IF #Stored = 0 THEN RETURN; END_IF;
    "FRK_PersistImages".D007.Rows[14] := "FRK_ConfigStore".Rows[#Stored];
    #Stored := "FRK_ConfigFind"(Scope := 'StationB.Satellite.Cell.Gate', Key := 'timeout', ModelCode := 'MODEL_B');
    IF #Stored = 0 THEN RETURN; END_IF;
    "FRK_PersistImages".D007.Rows[15] := "FRK_ConfigStore".Rows[#Stored];
    #Stored := "FRK_ConfigFind"(Scope := 'StationB.Satellite.Cell.Gate', Key := 'preset', ModelCode := 'MODEL_B');
    IF #Stored = 0 THEN RETURN; END_IF;
    "FRK_PersistImages".D007.Rows[16] := "FRK_ConfigStore".Rows[#Stored];
    #Stored := "FRK_ConfigFind"(Scope := 'StationB.Satellite.Inner', Key := 'timeout', ModelCode := 'MODEL_B');
    IF #Stored = 0 THEN RETURN; END_IF;
    "FRK_PersistImages".D007.Rows[17] := "FRK_ConfigStore".Rows[#Stored];
    #Stored := "FRK_ConfigFind"(Scope := 'StationB.Satellite.Inner', Key := 'preset', ModelCode := 'MODEL_B');
    IF #Stored = 0 THEN RETURN; END_IF;
    "FRK_PersistImages".D007.Rows[18] := "FRK_ConfigStore".Rows[#Stored];
    #Stored := "FRK_ConfigFind"(Scope := 'StationB.Satellite.Inner.Cell', Key := 'timeout', ModelCode := 'MODEL_B');
    IF #Stored = 0 THEN RETURN; END_IF;
    "FRK_PersistImages".D007.Rows[19] := "FRK_ConfigStore".Rows[#Stored];
    #Stored := "FRK_ConfigFind"(Scope := 'StationB.Satellite.Inner.Cell', Key := 'preset', ModelCode := 'MODEL_B');
    IF #Stored = 0 THEN RETURN; END_IF;
    "FRK_PersistImages".D007.Rows[20] := "FRK_ConfigStore".Rows[#Stored];
    #Stored := "FRK_ConfigFind"(Scope := 'StationB.Satellite.Inner.Cell.Clamp', Key := 'timeout', ModelCode := 'MODEL_B');
    IF #Stored = 0 THEN RETURN; END_IF;
    "FRK_PersistImages".D007.Rows[21] := "FRK_ConfigStore".Rows[#Stored];
    #Stored := "FRK_ConfigFind"(Scope := 'StationB.Satellite.Inner.Cell.Clamp', Key := 'preset', ModelCode := 'MODEL_B');
    IF #Stored = 0 THEN RETURN; END_IF;
    "FRK_PersistImages".D007.Rows[22] := "FRK_ConfigStore".Rows[#Stored];
    #Stored := "FRK_ConfigFind"(Scope := 'StationB.Satellite.Inner.Cell.Gate', Key := 'timeout', ModelCode := 'MODEL_B');
    IF #Stored = 0 THEN RETURN; END_IF;
    "FRK_PersistImages".D007.Rows[23] := "FRK_ConfigStore".Rows[#Stored];
    #Stored := "FRK_ConfigFind"(Scope := 'StationB.Satellite.Inner.Cell.Gate', Key := 'preset', ModelCode := 'MODEL_B');
    IF #Stored = 0 THEN RETURN; END_IF;
    "FRK_PersistImages".D007.Rows[24] := "FRK_ConfigStore".Rows[#Stored];
    FOR #Index := 0 TO 11401 DO "FRK_PersistBuffers".D007Data[#Index] := BYTE#0; END_FOR;
    #Position := 24;
    #NativeResult := Serialize(SRC_VARIABLE := "FRK_PersistImages".D007, DEST_ARRAY => "FRK_PersistBuffers".D007Data, POS := #Position);
    IF #NativeResult <> 0 OR #Position < 24 OR #Position > 11402 THEN RETURN; END_IF;
    #Length := #Position - 24;
    #FRK_DocCapture_D007 := TRUE;
END_FUNCTION
FUNCTION "FRK_DocApply_D007" : Bool
{ S7_Optimized_Access := 'TRUE' }
VERSION : 0.1
VAR_TEMP
    Index : Int;
    Stored : Int;
    Position : DInt;
    NativeResult : Int;
    Ok : Bool;
END_VAR
BEGIN
    #FRK_DocApply_D007 := FALSE;
    #Position := 24;
    #NativeResult := Deserialize(SRC_ARRAY := "FRK_PersistBuffers".D007Data, DEST_VARIABLE => "FRK_PersistImages".D007, POS := #Position);
    IF #NativeResult <> 0 OR #Position <> 24 + UDINT_TO_DINT("FRK_PersistConsumers".Rows[7].Result.Length) THEN RETURN; END_IF;
    IF "FRK_PersistImages".D007.SchemaVersion <> 1 OR "FRK_PersistImages".D007.Scope <> 'StationB' THEN RETURN; END_IF;
    IF "FRK_PersistImages".D007.Kind <> 0 OR "FRK_PersistImages".D007.ModelCode <> 'MODEL_B' OR "FRK_PersistImages".D007.Count <> 24 THEN RETURN; END_IF;
    IF "FRK_PersistImages".D007.ActiveModel <> 'MODEL_A' AND "FRK_PersistImages".D007.ActiveModel <> 'MODEL_B' THEN RETURN; END_IF;
    IF NOT "FRK_PersistImages".D007.Rows[1].Used OR "FRK_PersistImages".D007.Rows[1].SchemaVersion <> 4 OR "FRK_PersistImages".D007.Rows[1].ModelCode <> 'MODEL_B' OR "FRK_PersistImages".D007.Rows[1].Record.Scope <> 'StationB' OR "FRK_PersistImages".D007.Rows[1].Record.WriteKey <> 'timeout' OR "FRK_PersistImages".D007.Rows[1].Record.Revision <> 1 OR "FRK_PersistImages".D007.Rows[1].Record.Kind <> 0 OR "FRK_PersistImages".D007.Rows[1].Record.ValueType <> 3 THEN RETURN; END_IF;
    #Ok := "FRK_ConfigDecode"(Text := STRING_TO_WSTRING("FRK_PersistImages".D007.Rows[1].Record.ValueText), Storage := 7, Minimum := 1.0, Maximum := 60000.0, MaxLength := 0, Value := "FRK_ConfigScratch".Value);
    IF NOT #Ok THEN RETURN; END_IF;
    IF NOT "FRK_PersistImages".D007.Rows[2].Used OR "FRK_PersistImages".D007.Rows[2].SchemaVersion <> 4 OR "FRK_PersistImages".D007.Rows[2].ModelCode <> 'MODEL_B' OR "FRK_PersistImages".D007.Rows[2].Record.Scope <> 'StationB' OR "FRK_PersistImages".D007.Rows[2].Record.WriteKey <> 'preset' OR "FRK_PersistImages".D007.Rows[2].Record.Revision <> 2 OR "FRK_PersistImages".D007.Rows[2].Record.Kind <> 0 OR "FRK_PersistImages".D007.Rows[2].Record.ValueType <> 0 THEN RETURN; END_IF;
    #Ok := "FRK_ConfigDecode"(Text := STRING_TO_WSTRING("FRK_PersistImages".D007.Rows[2].Record.ValueText), Storage := 3, Minimum := 0.0, Maximum := 1000.0, MaxLength := 0, Value := "FRK_ConfigScratch".Value);
    IF NOT #Ok THEN RETURN; END_IF;
    IF NOT "FRK_PersistImages".D007.Rows[3].Used OR "FRK_PersistImages".D007.Rows[3].SchemaVersion <> 4 OR "FRK_PersistImages".D007.Rows[3].ModelCode <> 'MODEL_B' OR "FRK_PersistImages".D007.Rows[3].Record.Scope <> 'StationB.Cell' OR "FRK_PersistImages".D007.Rows[3].Record.WriteKey <> 'timeout' OR "FRK_PersistImages".D007.Rows[3].Record.Revision <> 1 OR "FRK_PersistImages".D007.Rows[3].Record.Kind <> 0 OR "FRK_PersistImages".D007.Rows[3].Record.ValueType <> 3 THEN RETURN; END_IF;
    #Ok := "FRK_ConfigDecode"(Text := STRING_TO_WSTRING("FRK_PersistImages".D007.Rows[3].Record.ValueText), Storage := 7, Minimum := 1.0, Maximum := 60000.0, MaxLength := 0, Value := "FRK_ConfigScratch".Value);
    IF NOT #Ok THEN RETURN; END_IF;
    IF NOT "FRK_PersistImages".D007.Rows[4].Used OR "FRK_PersistImages".D007.Rows[4].SchemaVersion <> 4 OR "FRK_PersistImages".D007.Rows[4].ModelCode <> 'MODEL_B' OR "FRK_PersistImages".D007.Rows[4].Record.Scope <> 'StationB.Cell' OR "FRK_PersistImages".D007.Rows[4].Record.WriteKey <> 'preset' OR "FRK_PersistImages".D007.Rows[4].Record.Revision <> 2 OR "FRK_PersistImages".D007.Rows[4].Record.Kind <> 0 OR "FRK_PersistImages".D007.Rows[4].Record.ValueType <> 0 THEN RETURN; END_IF;
    #Ok := "FRK_ConfigDecode"(Text := STRING_TO_WSTRING("FRK_PersistImages".D007.Rows[4].Record.ValueText), Storage := 3, Minimum := 0.0, Maximum := 1000.0, MaxLength := 0, Value := "FRK_ConfigScratch".Value);
    IF NOT #Ok THEN RETURN; END_IF;
    IF NOT "FRK_PersistImages".D007.Rows[5].Used OR "FRK_PersistImages".D007.Rows[5].SchemaVersion <> 4 OR "FRK_PersistImages".D007.Rows[5].ModelCode <> 'MODEL_B' OR "FRK_PersistImages".D007.Rows[5].Record.Scope <> 'StationB.Cell.Clamp' OR "FRK_PersistImages".D007.Rows[5].Record.WriteKey <> 'timeout' OR "FRK_PersistImages".D007.Rows[5].Record.Revision <> 1 OR "FRK_PersistImages".D007.Rows[5].Record.Kind <> 0 OR "FRK_PersistImages".D007.Rows[5].Record.ValueType <> 3 THEN RETURN; END_IF;
    #Ok := "FRK_ConfigDecode"(Text := STRING_TO_WSTRING("FRK_PersistImages".D007.Rows[5].Record.ValueText), Storage := 7, Minimum := 1.0, Maximum := 60000.0, MaxLength := 0, Value := "FRK_ConfigScratch".Value);
    IF NOT #Ok THEN RETURN; END_IF;
    IF NOT "FRK_PersistImages".D007.Rows[6].Used OR "FRK_PersistImages".D007.Rows[6].SchemaVersion <> 4 OR "FRK_PersistImages".D007.Rows[6].ModelCode <> 'MODEL_B' OR "FRK_PersistImages".D007.Rows[6].Record.Scope <> 'StationB.Cell.Clamp' OR "FRK_PersistImages".D007.Rows[6].Record.WriteKey <> 'preset' OR "FRK_PersistImages".D007.Rows[6].Record.Revision <> 2 OR "FRK_PersistImages".D007.Rows[6].Record.Kind <> 0 OR "FRK_PersistImages".D007.Rows[6].Record.ValueType <> 0 THEN RETURN; END_IF;
    #Ok := "FRK_ConfigDecode"(Text := STRING_TO_WSTRING("FRK_PersistImages".D007.Rows[6].Record.ValueText), Storage := 3, Minimum := 0.0, Maximum := 1000.0, MaxLength := 0, Value := "FRK_ConfigScratch".Value);
    IF NOT #Ok THEN RETURN; END_IF;
    IF NOT "FRK_PersistImages".D007.Rows[7].Used OR "FRK_PersistImages".D007.Rows[7].SchemaVersion <> 4 OR "FRK_PersistImages".D007.Rows[7].ModelCode <> 'MODEL_B' OR "FRK_PersistImages".D007.Rows[7].Record.Scope <> 'StationB.Cell.Gate' OR "FRK_PersistImages".D007.Rows[7].Record.WriteKey <> 'timeout' OR "FRK_PersistImages".D007.Rows[7].Record.Revision <> 1 OR "FRK_PersistImages".D007.Rows[7].Record.Kind <> 0 OR "FRK_PersistImages".D007.Rows[7].Record.ValueType <> 3 THEN RETURN; END_IF;
    #Ok := "FRK_ConfigDecode"(Text := STRING_TO_WSTRING("FRK_PersistImages".D007.Rows[7].Record.ValueText), Storage := 7, Minimum := 1.0, Maximum := 60000.0, MaxLength := 0, Value := "FRK_ConfigScratch".Value);
    IF NOT #Ok THEN RETURN; END_IF;
    IF NOT "FRK_PersistImages".D007.Rows[8].Used OR "FRK_PersistImages".D007.Rows[8].SchemaVersion <> 4 OR "FRK_PersistImages".D007.Rows[8].ModelCode <> 'MODEL_B' OR "FRK_PersistImages".D007.Rows[8].Record.Scope <> 'StationB.Cell.Gate' OR "FRK_PersistImages".D007.Rows[8].Record.WriteKey <> 'preset' OR "FRK_PersistImages".D007.Rows[8].Record.Revision <> 2 OR "FRK_PersistImages".D007.Rows[8].Record.Kind <> 0 OR "FRK_PersistImages".D007.Rows[8].Record.ValueType <> 0 THEN RETURN; END_IF;
    #Ok := "FRK_ConfigDecode"(Text := STRING_TO_WSTRING("FRK_PersistImages".D007.Rows[8].Record.ValueText), Storage := 3, Minimum := 0.0, Maximum := 1000.0, MaxLength := 0, Value := "FRK_ConfigScratch".Value);
    IF NOT #Ok THEN RETURN; END_IF;
    IF NOT "FRK_PersistImages".D007.Rows[9].Used OR "FRK_PersistImages".D007.Rows[9].SchemaVersion <> 4 OR "FRK_PersistImages".D007.Rows[9].ModelCode <> 'MODEL_B' OR "FRK_PersistImages".D007.Rows[9].Record.Scope <> 'StationB.Satellite' OR "FRK_PersistImages".D007.Rows[9].Record.WriteKey <> 'timeout' OR "FRK_PersistImages".D007.Rows[9].Record.Revision <> 1 OR "FRK_PersistImages".D007.Rows[9].Record.Kind <> 0 OR "FRK_PersistImages".D007.Rows[9].Record.ValueType <> 3 THEN RETURN; END_IF;
    #Ok := "FRK_ConfigDecode"(Text := STRING_TO_WSTRING("FRK_PersistImages".D007.Rows[9].Record.ValueText), Storage := 7, Minimum := 1.0, Maximum := 60000.0, MaxLength := 0, Value := "FRK_ConfigScratch".Value);
    IF NOT #Ok THEN RETURN; END_IF;
    IF NOT "FRK_PersistImages".D007.Rows[10].Used OR "FRK_PersistImages".D007.Rows[10].SchemaVersion <> 4 OR "FRK_PersistImages".D007.Rows[10].ModelCode <> 'MODEL_B' OR "FRK_PersistImages".D007.Rows[10].Record.Scope <> 'StationB.Satellite' OR "FRK_PersistImages".D007.Rows[10].Record.WriteKey <> 'preset' OR "FRK_PersistImages".D007.Rows[10].Record.Revision <> 2 OR "FRK_PersistImages".D007.Rows[10].Record.Kind <> 0 OR "FRK_PersistImages".D007.Rows[10].Record.ValueType <> 0 THEN RETURN; END_IF;
    #Ok := "FRK_ConfigDecode"(Text := STRING_TO_WSTRING("FRK_PersistImages".D007.Rows[10].Record.ValueText), Storage := 3, Minimum := 0.0, Maximum := 1000.0, MaxLength := 0, Value := "FRK_ConfigScratch".Value);
    IF NOT #Ok THEN RETURN; END_IF;
    IF NOT "FRK_PersistImages".D007.Rows[11].Used OR "FRK_PersistImages".D007.Rows[11].SchemaVersion <> 4 OR "FRK_PersistImages".D007.Rows[11].ModelCode <> 'MODEL_B' OR "FRK_PersistImages".D007.Rows[11].Record.Scope <> 'StationB.Satellite.Cell' OR "FRK_PersistImages".D007.Rows[11].Record.WriteKey <> 'timeout' OR "FRK_PersistImages".D007.Rows[11].Record.Revision <> 1 OR "FRK_PersistImages".D007.Rows[11].Record.Kind <> 0 OR "FRK_PersistImages".D007.Rows[11].Record.ValueType <> 3 THEN RETURN; END_IF;
    #Ok := "FRK_ConfigDecode"(Text := STRING_TO_WSTRING("FRK_PersistImages".D007.Rows[11].Record.ValueText), Storage := 7, Minimum := 1.0, Maximum := 60000.0, MaxLength := 0, Value := "FRK_ConfigScratch".Value);
    IF NOT #Ok THEN RETURN; END_IF;
    IF NOT "FRK_PersistImages".D007.Rows[12].Used OR "FRK_PersistImages".D007.Rows[12].SchemaVersion <> 4 OR "FRK_PersistImages".D007.Rows[12].ModelCode <> 'MODEL_B' OR "FRK_PersistImages".D007.Rows[12].Record.Scope <> 'StationB.Satellite.Cell' OR "FRK_PersistImages".D007.Rows[12].Record.WriteKey <> 'preset' OR "FRK_PersistImages".D007.Rows[12].Record.Revision <> 2 OR "FRK_PersistImages".D007.Rows[12].Record.Kind <> 0 OR "FRK_PersistImages".D007.Rows[12].Record.ValueType <> 0 THEN RETURN; END_IF;
    #Ok := "FRK_ConfigDecode"(Text := STRING_TO_WSTRING("FRK_PersistImages".D007.Rows[12].Record.ValueText), Storage := 3, Minimum := 0.0, Maximum := 1000.0, MaxLength := 0, Value := "FRK_ConfigScratch".Value);
    IF NOT #Ok THEN RETURN; END_IF;
    IF NOT "FRK_PersistImages".D007.Rows[13].Used OR "FRK_PersistImages".D007.Rows[13].SchemaVersion <> 4 OR "FRK_PersistImages".D007.Rows[13].ModelCode <> 'MODEL_B' OR "FRK_PersistImages".D007.Rows[13].Record.Scope <> 'StationB.Satellite.Cell.Clamp' OR "FRK_PersistImages".D007.Rows[13].Record.WriteKey <> 'timeout' OR "FRK_PersistImages".D007.Rows[13].Record.Revision <> 1 OR "FRK_PersistImages".D007.Rows[13].Record.Kind <> 0 OR "FRK_PersistImages".D007.Rows[13].Record.ValueType <> 3 THEN RETURN; END_IF;
    #Ok := "FRK_ConfigDecode"(Text := STRING_TO_WSTRING("FRK_PersistImages".D007.Rows[13].Record.ValueText), Storage := 7, Minimum := 1.0, Maximum := 60000.0, MaxLength := 0, Value := "FRK_ConfigScratch".Value);
    IF NOT #Ok THEN RETURN; END_IF;
    IF NOT "FRK_PersistImages".D007.Rows[14].Used OR "FRK_PersistImages".D007.Rows[14].SchemaVersion <> 4 OR "FRK_PersistImages".D007.Rows[14].ModelCode <> 'MODEL_B' OR "FRK_PersistImages".D007.Rows[14].Record.Scope <> 'StationB.Satellite.Cell.Clamp' OR "FRK_PersistImages".D007.Rows[14].Record.WriteKey <> 'preset' OR "FRK_PersistImages".D007.Rows[14].Record.Revision <> 2 OR "FRK_PersistImages".D007.Rows[14].Record.Kind <> 0 OR "FRK_PersistImages".D007.Rows[14].Record.ValueType <> 0 THEN RETURN; END_IF;
    #Ok := "FRK_ConfigDecode"(Text := STRING_TO_WSTRING("FRK_PersistImages".D007.Rows[14].Record.ValueText), Storage := 3, Minimum := 0.0, Maximum := 1000.0, MaxLength := 0, Value := "FRK_ConfigScratch".Value);
    IF NOT #Ok THEN RETURN; END_IF;
    IF NOT "FRK_PersistImages".D007.Rows[15].Used OR "FRK_PersistImages".D007.Rows[15].SchemaVersion <> 4 OR "FRK_PersistImages".D007.Rows[15].ModelCode <> 'MODEL_B' OR "FRK_PersistImages".D007.Rows[15].Record.Scope <> 'StationB.Satellite.Cell.Gate' OR "FRK_PersistImages".D007.Rows[15].Record.WriteKey <> 'timeout' OR "FRK_PersistImages".D007.Rows[15].Record.Revision <> 1 OR "FRK_PersistImages".D007.Rows[15].Record.Kind <> 0 OR "FRK_PersistImages".D007.Rows[15].Record.ValueType <> 3 THEN RETURN; END_IF;
    #Ok := "FRK_ConfigDecode"(Text := STRING_TO_WSTRING("FRK_PersistImages".D007.Rows[15].Record.ValueText), Storage := 7, Minimum := 1.0, Maximum := 60000.0, MaxLength := 0, Value := "FRK_ConfigScratch".Value);
    IF NOT #Ok THEN RETURN; END_IF;
    IF NOT "FRK_PersistImages".D007.Rows[16].Used OR "FRK_PersistImages".D007.Rows[16].SchemaVersion <> 4 OR "FRK_PersistImages".D007.Rows[16].ModelCode <> 'MODEL_B' OR "FRK_PersistImages".D007.Rows[16].Record.Scope <> 'StationB.Satellite.Cell.Gate' OR "FRK_PersistImages".D007.Rows[16].Record.WriteKey <> 'preset' OR "FRK_PersistImages".D007.Rows[16].Record.Revision <> 2 OR "FRK_PersistImages".D007.Rows[16].Record.Kind <> 0 OR "FRK_PersistImages".D007.Rows[16].Record.ValueType <> 0 THEN RETURN; END_IF;
    #Ok := "FRK_ConfigDecode"(Text := STRING_TO_WSTRING("FRK_PersistImages".D007.Rows[16].Record.ValueText), Storage := 3, Minimum := 0.0, Maximum := 1000.0, MaxLength := 0, Value := "FRK_ConfigScratch".Value);
    IF NOT #Ok THEN RETURN; END_IF;
    IF NOT "FRK_PersistImages".D007.Rows[17].Used OR "FRK_PersistImages".D007.Rows[17].SchemaVersion <> 4 OR "FRK_PersistImages".D007.Rows[17].ModelCode <> 'MODEL_B' OR "FRK_PersistImages".D007.Rows[17].Record.Scope <> 'StationB.Satellite.Inner' OR "FRK_PersistImages".D007.Rows[17].Record.WriteKey <> 'timeout' OR "FRK_PersistImages".D007.Rows[17].Record.Revision <> 1 OR "FRK_PersistImages".D007.Rows[17].Record.Kind <> 0 OR "FRK_PersistImages".D007.Rows[17].Record.ValueType <> 3 THEN RETURN; END_IF;
    #Ok := "FRK_ConfigDecode"(Text := STRING_TO_WSTRING("FRK_PersistImages".D007.Rows[17].Record.ValueText), Storage := 7, Minimum := 1.0, Maximum := 60000.0, MaxLength := 0, Value := "FRK_ConfigScratch".Value);
    IF NOT #Ok THEN RETURN; END_IF;
    IF NOT "FRK_PersistImages".D007.Rows[18].Used OR "FRK_PersistImages".D007.Rows[18].SchemaVersion <> 4 OR "FRK_PersistImages".D007.Rows[18].ModelCode <> 'MODEL_B' OR "FRK_PersistImages".D007.Rows[18].Record.Scope <> 'StationB.Satellite.Inner' OR "FRK_PersistImages".D007.Rows[18].Record.WriteKey <> 'preset' OR "FRK_PersistImages".D007.Rows[18].Record.Revision <> 2 OR "FRK_PersistImages".D007.Rows[18].Record.Kind <> 0 OR "FRK_PersistImages".D007.Rows[18].Record.ValueType <> 0 THEN RETURN; END_IF;
    #Ok := "FRK_ConfigDecode"(Text := STRING_TO_WSTRING("FRK_PersistImages".D007.Rows[18].Record.ValueText), Storage := 3, Minimum := 0.0, Maximum := 1000.0, MaxLength := 0, Value := "FRK_ConfigScratch".Value);
    IF NOT #Ok THEN RETURN; END_IF;
    IF NOT "FRK_PersistImages".D007.Rows[19].Used OR "FRK_PersistImages".D007.Rows[19].SchemaVersion <> 4 OR "FRK_PersistImages".D007.Rows[19].ModelCode <> 'MODEL_B' OR "FRK_PersistImages".D007.Rows[19].Record.Scope <> 'StationB.Satellite.Inner.Cell' OR "FRK_PersistImages".D007.Rows[19].Record.WriteKey <> 'timeout' OR "FRK_PersistImages".D007.Rows[19].Record.Revision <> 1 OR "FRK_PersistImages".D007.Rows[19].Record.Kind <> 0 OR "FRK_PersistImages".D007.Rows[19].Record.ValueType <> 3 THEN RETURN; END_IF;
    #Ok := "FRK_ConfigDecode"(Text := STRING_TO_WSTRING("FRK_PersistImages".D007.Rows[19].Record.ValueText), Storage := 7, Minimum := 1.0, Maximum := 60000.0, MaxLength := 0, Value := "FRK_ConfigScratch".Value);
    IF NOT #Ok THEN RETURN; END_IF;
    IF NOT "FRK_PersistImages".D007.Rows[20].Used OR "FRK_PersistImages".D007.Rows[20].SchemaVersion <> 4 OR "FRK_PersistImages".D007.Rows[20].ModelCode <> 'MODEL_B' OR "FRK_PersistImages".D007.Rows[20].Record.Scope <> 'StationB.Satellite.Inner.Cell' OR "FRK_PersistImages".D007.Rows[20].Record.WriteKey <> 'preset' OR "FRK_PersistImages".D007.Rows[20].Record.Revision <> 2 OR "FRK_PersistImages".D007.Rows[20].Record.Kind <> 0 OR "FRK_PersistImages".D007.Rows[20].Record.ValueType <> 0 THEN RETURN; END_IF;
    #Ok := "FRK_ConfigDecode"(Text := STRING_TO_WSTRING("FRK_PersistImages".D007.Rows[20].Record.ValueText), Storage := 3, Minimum := 0.0, Maximum := 1000.0, MaxLength := 0, Value := "FRK_ConfigScratch".Value);
    IF NOT #Ok THEN RETURN; END_IF;
    IF NOT "FRK_PersistImages".D007.Rows[21].Used OR "FRK_PersistImages".D007.Rows[21].SchemaVersion <> 4 OR "FRK_PersistImages".D007.Rows[21].ModelCode <> 'MODEL_B' OR "FRK_PersistImages".D007.Rows[21].Record.Scope <> 'StationB.Satellite.Inner.Cell.Clamp' OR "FRK_PersistImages".D007.Rows[21].Record.WriteKey <> 'timeout' OR "FRK_PersistImages".D007.Rows[21].Record.Revision <> 1 OR "FRK_PersistImages".D007.Rows[21].Record.Kind <> 0 OR "FRK_PersistImages".D007.Rows[21].Record.ValueType <> 3 THEN RETURN; END_IF;
    #Ok := "FRK_ConfigDecode"(Text := STRING_TO_WSTRING("FRK_PersistImages".D007.Rows[21].Record.ValueText), Storage := 7, Minimum := 1.0, Maximum := 60000.0, MaxLength := 0, Value := "FRK_ConfigScratch".Value);
    IF NOT #Ok THEN RETURN; END_IF;
    IF NOT "FRK_PersistImages".D007.Rows[22].Used OR "FRK_PersistImages".D007.Rows[22].SchemaVersion <> 4 OR "FRK_PersistImages".D007.Rows[22].ModelCode <> 'MODEL_B' OR "FRK_PersistImages".D007.Rows[22].Record.Scope <> 'StationB.Satellite.Inner.Cell.Clamp' OR "FRK_PersistImages".D007.Rows[22].Record.WriteKey <> 'preset' OR "FRK_PersistImages".D007.Rows[22].Record.Revision <> 2 OR "FRK_PersistImages".D007.Rows[22].Record.Kind <> 0 OR "FRK_PersistImages".D007.Rows[22].Record.ValueType <> 0 THEN RETURN; END_IF;
    #Ok := "FRK_ConfigDecode"(Text := STRING_TO_WSTRING("FRK_PersistImages".D007.Rows[22].Record.ValueText), Storage := 3, Minimum := 0.0, Maximum := 1000.0, MaxLength := 0, Value := "FRK_ConfigScratch".Value);
    IF NOT #Ok THEN RETURN; END_IF;
    IF NOT "FRK_PersistImages".D007.Rows[23].Used OR "FRK_PersistImages".D007.Rows[23].SchemaVersion <> 4 OR "FRK_PersistImages".D007.Rows[23].ModelCode <> 'MODEL_B' OR "FRK_PersistImages".D007.Rows[23].Record.Scope <> 'StationB.Satellite.Inner.Cell.Gate' OR "FRK_PersistImages".D007.Rows[23].Record.WriteKey <> 'timeout' OR "FRK_PersistImages".D007.Rows[23].Record.Revision <> 1 OR "FRK_PersistImages".D007.Rows[23].Record.Kind <> 0 OR "FRK_PersistImages".D007.Rows[23].Record.ValueType <> 3 THEN RETURN; END_IF;
    #Ok := "FRK_ConfigDecode"(Text := STRING_TO_WSTRING("FRK_PersistImages".D007.Rows[23].Record.ValueText), Storage := 7, Minimum := 1.0, Maximum := 60000.0, MaxLength := 0, Value := "FRK_ConfigScratch".Value);
    IF NOT #Ok THEN RETURN; END_IF;
    IF NOT "FRK_PersistImages".D007.Rows[24].Used OR "FRK_PersistImages".D007.Rows[24].SchemaVersion <> 4 OR "FRK_PersistImages".D007.Rows[24].ModelCode <> 'MODEL_B' OR "FRK_PersistImages".D007.Rows[24].Record.Scope <> 'StationB.Satellite.Inner.Cell.Gate' OR "FRK_PersistImages".D007.Rows[24].Record.WriteKey <> 'preset' OR "FRK_PersistImages".D007.Rows[24].Record.Revision <> 2 OR "FRK_PersistImages".D007.Rows[24].Record.Kind <> 0 OR "FRK_PersistImages".D007.Rows[24].Record.ValueType <> 0 THEN RETURN; END_IF;
    #Ok := "FRK_ConfigDecode"(Text := STRING_TO_WSTRING("FRK_PersistImages".D007.Rows[24].Record.ValueText), Storage := 3, Minimum := 0.0, Maximum := 1000.0, MaxLength := 0, Value := "FRK_ConfigScratch".Value);
    IF NOT #Ok THEN RETURN; END_IF;
    #Stored := "FRK_ConfigFind"(Scope := 'StationB', Key := 'timeout', ModelCode := 'MODEL_B');
    IF #Stored = 0 THEN
        FOR #Stored := 1 TO 108 DO IF NOT "FRK_ConfigStore".Rows[#Stored].Used THEN EXIT; END_IF; END_FOR;
    END_IF;
    IF #Stored < 1 OR #Stored > 108 THEN RETURN; END_IF;
    "FRK_ConfigStore".Rows[#Stored] := "FRK_PersistImages".D007.Rows[1];
    #Stored := "FRK_ConfigFind"(Scope := 'StationB', Key := 'preset', ModelCode := 'MODEL_B');
    IF #Stored = 0 THEN
        FOR #Stored := 1 TO 108 DO IF NOT "FRK_ConfigStore".Rows[#Stored].Used THEN EXIT; END_IF; END_FOR;
    END_IF;
    IF #Stored < 1 OR #Stored > 108 THEN RETURN; END_IF;
    "FRK_ConfigStore".Rows[#Stored] := "FRK_PersistImages".D007.Rows[2];
    #Stored := "FRK_ConfigFind"(Scope := 'StationB.Cell', Key := 'timeout', ModelCode := 'MODEL_B');
    IF #Stored = 0 THEN
        FOR #Stored := 1 TO 108 DO IF NOT "FRK_ConfigStore".Rows[#Stored].Used THEN EXIT; END_IF; END_FOR;
    END_IF;
    IF #Stored < 1 OR #Stored > 108 THEN RETURN; END_IF;
    "FRK_ConfigStore".Rows[#Stored] := "FRK_PersistImages".D007.Rows[3];
    #Stored := "FRK_ConfigFind"(Scope := 'StationB.Cell', Key := 'preset', ModelCode := 'MODEL_B');
    IF #Stored = 0 THEN
        FOR #Stored := 1 TO 108 DO IF NOT "FRK_ConfigStore".Rows[#Stored].Used THEN EXIT; END_IF; END_FOR;
    END_IF;
    IF #Stored < 1 OR #Stored > 108 THEN RETURN; END_IF;
    "FRK_ConfigStore".Rows[#Stored] := "FRK_PersistImages".D007.Rows[4];
    #Stored := "FRK_ConfigFind"(Scope := 'StationB.Cell.Clamp', Key := 'timeout', ModelCode := 'MODEL_B');
    IF #Stored = 0 THEN
        FOR #Stored := 1 TO 108 DO IF NOT "FRK_ConfigStore".Rows[#Stored].Used THEN EXIT; END_IF; END_FOR;
    END_IF;
    IF #Stored < 1 OR #Stored > 108 THEN RETURN; END_IF;
    "FRK_ConfigStore".Rows[#Stored] := "FRK_PersistImages".D007.Rows[5];
    #Stored := "FRK_ConfigFind"(Scope := 'StationB.Cell.Clamp', Key := 'preset', ModelCode := 'MODEL_B');
    IF #Stored = 0 THEN
        FOR #Stored := 1 TO 108 DO IF NOT "FRK_ConfigStore".Rows[#Stored].Used THEN EXIT; END_IF; END_FOR;
    END_IF;
    IF #Stored < 1 OR #Stored > 108 THEN RETURN; END_IF;
    "FRK_ConfigStore".Rows[#Stored] := "FRK_PersistImages".D007.Rows[6];
    #Stored := "FRK_ConfigFind"(Scope := 'StationB.Cell.Gate', Key := 'timeout', ModelCode := 'MODEL_B');
    IF #Stored = 0 THEN
        FOR #Stored := 1 TO 108 DO IF NOT "FRK_ConfigStore".Rows[#Stored].Used THEN EXIT; END_IF; END_FOR;
    END_IF;
    IF #Stored < 1 OR #Stored > 108 THEN RETURN; END_IF;
    "FRK_ConfigStore".Rows[#Stored] := "FRK_PersistImages".D007.Rows[7];
    #Stored := "FRK_ConfigFind"(Scope := 'StationB.Cell.Gate', Key := 'preset', ModelCode := 'MODEL_B');
    IF #Stored = 0 THEN
        FOR #Stored := 1 TO 108 DO IF NOT "FRK_ConfigStore".Rows[#Stored].Used THEN EXIT; END_IF; END_FOR;
    END_IF;
    IF #Stored < 1 OR #Stored > 108 THEN RETURN; END_IF;
    "FRK_ConfigStore".Rows[#Stored] := "FRK_PersistImages".D007.Rows[8];
    #Stored := "FRK_ConfigFind"(Scope := 'StationB.Satellite', Key := 'timeout', ModelCode := 'MODEL_B');
    IF #Stored = 0 THEN
        FOR #Stored := 1 TO 108 DO IF NOT "FRK_ConfigStore".Rows[#Stored].Used THEN EXIT; END_IF; END_FOR;
    END_IF;
    IF #Stored < 1 OR #Stored > 108 THEN RETURN; END_IF;
    "FRK_ConfigStore".Rows[#Stored] := "FRK_PersistImages".D007.Rows[9];
    #Stored := "FRK_ConfigFind"(Scope := 'StationB.Satellite', Key := 'preset', ModelCode := 'MODEL_B');
    IF #Stored = 0 THEN
        FOR #Stored := 1 TO 108 DO IF NOT "FRK_ConfigStore".Rows[#Stored].Used THEN EXIT; END_IF; END_FOR;
    END_IF;
    IF #Stored < 1 OR #Stored > 108 THEN RETURN; END_IF;
    "FRK_ConfigStore".Rows[#Stored] := "FRK_PersistImages".D007.Rows[10];
    #Stored := "FRK_ConfigFind"(Scope := 'StationB.Satellite.Cell', Key := 'timeout', ModelCode := 'MODEL_B');
    IF #Stored = 0 THEN
        FOR #Stored := 1 TO 108 DO IF NOT "FRK_ConfigStore".Rows[#Stored].Used THEN EXIT; END_IF; END_FOR;
    END_IF;
    IF #Stored < 1 OR #Stored > 108 THEN RETURN; END_IF;
    "FRK_ConfigStore".Rows[#Stored] := "FRK_PersistImages".D007.Rows[11];
    #Stored := "FRK_ConfigFind"(Scope := 'StationB.Satellite.Cell', Key := 'preset', ModelCode := 'MODEL_B');
    IF #Stored = 0 THEN
        FOR #Stored := 1 TO 108 DO IF NOT "FRK_ConfigStore".Rows[#Stored].Used THEN EXIT; END_IF; END_FOR;
    END_IF;
    IF #Stored < 1 OR #Stored > 108 THEN RETURN; END_IF;
    "FRK_ConfigStore".Rows[#Stored] := "FRK_PersistImages".D007.Rows[12];
    #Stored := "FRK_ConfigFind"(Scope := 'StationB.Satellite.Cell.Clamp', Key := 'timeout', ModelCode := 'MODEL_B');
    IF #Stored = 0 THEN
        FOR #Stored := 1 TO 108 DO IF NOT "FRK_ConfigStore".Rows[#Stored].Used THEN EXIT; END_IF; END_FOR;
    END_IF;
    IF #Stored < 1 OR #Stored > 108 THEN RETURN; END_IF;
    "FRK_ConfigStore".Rows[#Stored] := "FRK_PersistImages".D007.Rows[13];
    #Stored := "FRK_ConfigFind"(Scope := 'StationB.Satellite.Cell.Clamp', Key := 'preset', ModelCode := 'MODEL_B');
    IF #Stored = 0 THEN
        FOR #Stored := 1 TO 108 DO IF NOT "FRK_ConfigStore".Rows[#Stored].Used THEN EXIT; END_IF; END_FOR;
    END_IF;
    IF #Stored < 1 OR #Stored > 108 THEN RETURN; END_IF;
    "FRK_ConfigStore".Rows[#Stored] := "FRK_PersistImages".D007.Rows[14];
    #Stored := "FRK_ConfigFind"(Scope := 'StationB.Satellite.Cell.Gate', Key := 'timeout', ModelCode := 'MODEL_B');
    IF #Stored = 0 THEN
        FOR #Stored := 1 TO 108 DO IF NOT "FRK_ConfigStore".Rows[#Stored].Used THEN EXIT; END_IF; END_FOR;
    END_IF;
    IF #Stored < 1 OR #Stored > 108 THEN RETURN; END_IF;
    "FRK_ConfigStore".Rows[#Stored] := "FRK_PersistImages".D007.Rows[15];
    #Stored := "FRK_ConfigFind"(Scope := 'StationB.Satellite.Cell.Gate', Key := 'preset', ModelCode := 'MODEL_B');
    IF #Stored = 0 THEN
        FOR #Stored := 1 TO 108 DO IF NOT "FRK_ConfigStore".Rows[#Stored].Used THEN EXIT; END_IF; END_FOR;
    END_IF;
    IF #Stored < 1 OR #Stored > 108 THEN RETURN; END_IF;
    "FRK_ConfigStore".Rows[#Stored] := "FRK_PersistImages".D007.Rows[16];
